(* IEC 61131-3 sources: daoli-st-library/DL_Device (part 33) *)

(* ---- FB_DL_ThreePointValve.st ---- *)
(*==============================================================================
 * 组件名称 (Component)  : FB_DL_ThreePointValve
 * 所属子库 (Sublibrary) : DL_Device
 * 当前版本 (Version)    : 1.0.1
 * 兼容性   (Platform)   : CODESYS 3.5 / TwinCAT 3 / 汇川 InoProShop / Machine Expert
 *                         仅依赖 Standard.library（TON / R_TRIG），零厂商方言
 * 分类     (Category)   : 设备执行器功能块（Function Block，实现 I_DL_MotorizedValve）
 * 功能简述 (Function)   : 三点浮点式电动调节阀控制器。开/关双脉冲输出；
 *                         行程时间积分自动估算开度（TON 计时段 ET 折算，
 *                         量纲推导见段 4 注释）；全开/全关限位双保险保护
 *                         （限位锚定 + 无限位端点拒绝）；限位互斥与估算-
 *                         限位一致性监视；双向指令互斥；首扫按限位状态
 *                         推断初值（R19 范式，bTrack 强制重同步）；状态机
 *                         E_DL_MotorValveState + CASE + ELSE 兜底。
 * 接口实现 (Implements) : I_DL_MotorizedValve。接口 OUT 列同名成员
 *                         （eState/fPosEstimate/bLimOpen/bLimClosed/
 *                         bFault/uErrorId）按 R22 以只读 PROPERTY GET 承载
 *                         （内部镜像同源；fPosEstimate 为 OUT 引脚、
 *                         bLimOpen/bLimClosed 为 IN 引脚与接口属性双形式
 *                         暴露，沿用库级既有先例），非接口成员 bOpenPulse/
 *                         bClosePulse/bOpened/bClosed/uTravelCount 保留
 *                         VAR_OUTPUT；方法 CmdOpen/CmdClose/CmdStop/
 *                         CmdReset 全部在本文件尾部落地。
 * 开源溯源 (Origin)     : 来源标签 lbp-basic-process / lbp-device
 *                         （RAW_NOTES_R6 S-1 + S-5：三点浮点式电动阀的开/
 *                         关脉冲控制、行程时间开度积分估算、端点限位双
 *                         保险等行业公知工程惯例，公开教学资料，仅借鉴
 *                         通用工程语义；状态机、积分实现、故障码按本库
 *                         红线独立设计，clean-room 未复制源码）。
 * 红线自检 (Redline)    : R1 零全局变量表/外部变量引用 ✓｜R2 零物理 IO 地址 ✓
 *                         R3 纯 IEC 61131-3 ✓｜R4 防除零/防越界/浮点容差
 *                         比较 ✓｜R5 全变量中英双语同行注释 ✓
 *                         R6 ENUM+CASE+ELSE ✓｜R7 四个定时器/边缘实例主体
 *                         最前部无条件刷新 ✓
 * 公约遵循 (Convention) : 0.1/R19 本块为事件型 + 连续估算混合组件：开度
 *                         积分为连续量，设 bInit 首扫（初值 FALSE，同步后
 *                         置 TRUE），判据唯一合法范式 IF bTrack OR (NOT
 *                         bInit)；bTrack 引脚供上层运行中途强制重同步。
 *                         0.7 故障码段位 16#0003_xxxx：【故障级】0003_0270
 *                         行程估算失准 / 0003_0271 双限位冲突 / 0003_0272
 *                         非法状态，R15 锁存仅复位可清；【信息级】
 *                         0003_0110 端点指令拒绝 / 0003_0111 双向指令冲突
 *                         （瞬时型每拍重算，0.15；不进 bFault）。
 * 偏离留档 (Deviation)  : 依 R11 头注释留档，共 3 条：
 *                         ① 信息级码：规格原分配 0003_0107/0108，经与子库
 *                           VERSION.md 故障码表核对，R5 已占用 0102~0104，
 *                           且 0106~0109 已由本轮变频器/模拟量阀块顺延占用
 *                           （0105 经终审裁定空置：重启抑制拒绝统一沿用
 *                           DolMotor 既有语义码位 0208），依公约 0.7 冲突
 *                           顺延为 0003_0110/0111。
 *                         ② 开度积分：规格原文"每拍按 fDt 增量累加"需周期
 *                           时间注入或时钟基准（与公约 0.9 冲突）；本实现
 *                           改用 TON 计时段 ET 累计行程时间折算：
 *                           fPosEstimate = 锚点 + 100 × ET[ms] / 行程时间[ms]
 *                           （量纲推导：无量纲比值 × 100% = [%]），等价
 *                           消除逐拍折算误差且零时钟依赖。
 *                         ③ bOpened/bClosed 的估算近似判据取固定 1% 吸附带
 *                           （限位优先，无限位场景估算到端点 1% 带内即视为
 *                           确认），规格未定值，现场可按需整定行程时间。
 * 修订历史 (Revision)   :
 *   2026-11-15  v1.0.0  首版入库（R6 轮 · DL_Device 阀门/驱动族深化）
 *   2026-11-15  v1.0.1  终审注释级修订：头注释偏离①码位占位表述与终审裁定
 *                       对齐（0105 空置、重启抑制拒绝归一 DolMotor 0208）。
 *                       逻辑零变更。已知诊断口径观察项（不改码）：uTravelCount
 *                       在上电首扫若全关限位已压住会即计 +1（限位态计数），
 *                       与 R4 PwmDutyController 首周期计数偏差同类，±1 口径。
 *============================================================================*)
FUNCTION_BLOCK FB_DL_ThreePointValve IMPLEMENTS I_DL_MotorizedValve
VAR_INPUT
    bCmdOpen     : BOOL;            // 开阀指令（Open command），电平生效 / Open command, level effective
    bCmdClose    : BOOL;            // 关阀指令（Close command），电平生效；与开同拍为真 → 停止 + 信息级 / Close command, conflict with open stops with info code
    bLimOpen     : BOOL;            // 全开限位开关（Open limit switch），TRUE=已到全开端点 / Open limit switch, TRUE = at fully-open endpoint
    bLimClosed   : BOOL;            // 全关限位开关（Closed limit switch），TRUE=已到全关端点 / Closed limit switch, TRUE = at fully-closed endpoint
    tStrokeOpen  : TIME := T#60S;   // 全行程开启时间（Full open stroke time），现场实测注入 / Full-open stroke time, field-measured
    tStrokeClose : TIME := T#60S;   // 全行程关闭时间（Full close stroke time），现场实测注入 / Full-close stroke time, field-measured
    fEstimateTol : REAL := 10.0;    // 估算-限位一致性容差（Estimate tolerance）[%]，默认 10.0 / Estimate-vs-limit consistency tolerance [%]
    bEnable      : BOOL;            // 允许动作联锁（Motion interlock），TRUE=允许发脉冲 / Motion interlock, TRUE = pulses allowed
    bReset       : BOOL;            // 故障复位（Fault reset），上升沿生效 / Fault reset, rising edge effective
    bTrack       : BOOL;            // 跟踪重同步（Track resync），TRUE 拍按限位状态重推初值（R19）/ Track resync re-infers initial estimate from limits
END_VAR

VAR_OUTPUT
    bOpenPulse   : BOOL;            // 开阀脉冲输出（Open pulse output）/ Open pulse output
    bClosePulse  : BOOL;            // 关阀脉冲输出（Close pulse output）/ Close pulse output
    fPosEstimate : REAL;            // 估算开度（Estimated position）[%]，0~100，行程时间积分（R20：量纲 [%]）/ Estimated position [%], stroke-time integration
    bOpened      : BOOL;            // 全开确认（Fully opened），限位优先 / Fully opened, limit switch has priority
    bClosed      : BOOL;            // 全关确认（Fully closed），限位优先 / Fully closed, limit switch has priority
    uTravelCount : UDINT;           // 全行程计数（Travel count），全关确认沿 +1 / Travel count, incremented on closed-confirmation edge
END_VAR

VAR
    _eState        : E_DL_MotorValveState := E_DL_MotorValveState.eIdle; // 内部状态机步序（Internal state step），外部经属性只读 / Internal state, read-only via property
    _bInit         : BOOL := FALSE; // 首扫初始化标志（First-scan init flag），R19 范式判据成员 / R19 paradigm member
    _bFaultLatch   : BOOL;          // 故障锁存标志（Fault latch flag），仅复位清除 / Fault latch flag, cleared only by reset
    _uErrorIdInt   : UDINT;         // 故障级码内部寄存（Internal fault-code register）/ Internal fault-level code register
    _uInfoCode     : UDINT;         // 本拍信息级码（Info code this cycle），瞬时型每拍重算（0.15）/ Transient info code recomputed each cycle
    _fAnchor       : REAL := 50.0;  // 积分锚点（Integration anchor）[%]，脉冲静止期与估算值同步 / Integration anchor [%], synced with estimate when idle
    _fEstInt       : REAL := 50.0;  // 估算开度内部寄存（Internal estimate register）[%] / Internal estimate register [%]
    _bPendOpen     : BOOL;          // 方法开阀保持锁存（Method open hold latch）/ Method open hold latch
    _bPendClose    : BOOL;          // 方法关阀保持锁存（Method close hold latch）/ Method close hold latch
    _bPendStop     : BOOL;          // 方法停止请求（Method stop request），由 CmdStop 置位 / Method stop request set by CmdStop
    _bPendReset    : BOOL;          // 方法复位请求（Method reset request），由 CmdReset 置位 / Method reset request set by CmdReset
    _bOpenReq      : BOOL;          // 合成开阀指令（Merged open command），引脚 OR 方法锁存 / Merged open command, pin OR method latch
    _bCloseReq     : BOOL;          // 合成关阀指令（Merged close command），引脚 OR 方法锁存 / Merged close command, pin OR method latch
    _bConflict     : BOOL;          // 双向同拍冲突（Open/close conflict this cycle）/ Open-close conflict flag
    _bOpenAtEnd    : BOOL;          // 开端点到达（Open endpoint reached），限位或估算判据 / Open endpoint reached by limit or estimate
    _bCloseAtEnd   : BOOL;          // 关端点到达（Close endpoint reached），限位或估算判据 / Close endpoint reached by limit or estimate
    _fTolEff       : REAL := 10.0;  // 防御后一致性容差（Sanitized tolerance）[%] / Sanitized consistency tolerance
    _tStrokeOpenEff  : TIME := T#60S; // 防御后开启行程时间（Sanitized open stroke time），非正值回退默认 / Sanitized open stroke time, non-positive falls back
    _tStrokeCloseEff : TIME := T#60S; // 防御后关闭行程时间（Sanitized close stroke time），非正值回退默认 / Sanitized close stroke time, non-positive falls back
    _bClosedInt    : BOOL;          // 全关确认内部镜像（Internal closed-confirmation mirror），喂计数边缘实例 / Internal closed mirror feeding count edge
    _bLimOpenMir   : BOOL;          // 全开限位内部镜像（Internal open-limit mirror），供属性读取 / Internal open-limit mirror for property exposure
    _bLimClosedMir : BOOL;          // 全关限位内部镜像（Internal closed-limit mirror），供属性读取 / Internal closed-limit mirror for property exposure
    _fbTrigReset   : R_TRIG;        // 引脚复位上升沿（Pin reset edge）/ Pin reset rising edge
    _fbTrigTravel  : R_TRIG;        // 全关确认计数上升沿（Travel count edge）/ Rising edge on closed confirmation for counting
    _fbTonOpenET   : TON;           // 开阀计时段定时器（Open timing segment timer），ET 供积分折算 / Open segment timer, ET feeds integration
    _fbTonCloseET  : TON;           // 关阀计时段定时器（Close timing segment timer），ET 供积分折算 / Close segment timer, ET feeds integration
END_VAR

METHOD CmdOpen : BOOL
VAR_INPUT
END_VAR
IF _bFaultLatch OR (_eState = E_DL_MotorValveState.eFault) THEN
    CmdOpen := FALSE;         // 故障态拒绝（Rejected in fault state）
    _bPendClose := FALSE;     // 清反向残留锁存（Clear stale reverse latch）
ELSE
    _bPendOpen := TRUE;       // 登记开阀保持锁存（Register open hold latch）
    _bPendClose := FALSE;     // 互斥注销关阀锁存（Cancel opposite close latch）
    CmdOpen := TRUE;          // 受理成功（Accepted）
END_IF

(*------------------------------------------------------------------------------
 * 方法: CmdClose —— 关阀指令（受理为保持锁存）。故障态一律拒绝返回 FALSE。
 *      Method CmdClose - close command held as latch, rejected with FALSE in fault.
 *------------------------------------------------------------------------------*)
    END_METHOD

METHOD CmdClose : BOOL
VAR_INPUT
END_VAR
IF _bFaultLatch OR (_eState = E_DL_MotorValveState.eFault) THEN
    CmdClose := FALSE;        // 故障态拒绝（Rejected in fault state）
    _bPendOpen := FALSE;      // 清反向残留锁存（Clear stale reverse latch）
ELSE
    _bPendClose := TRUE;      // 登记关阀保持锁存（Register close hold latch）
    _bPendOpen := FALSE;      // 互斥注销开阀锁存（Cancel opposite open latch）
    CmdClose := TRUE;         // 受理成功（Accepted）
END_IF

(*------------------------------------------------------------------------------
 * 方法: CmdStop —— 双脉冲全断保持当前位置。无条件受理。
 *      Method CmdStop - both pulses off and hold position, unconditionally accepted.
 *------------------------------------------------------------------------------*)
    END_METHOD

METHOD CmdStop : BOOL
VAR_INPUT
END_VAR
_bPendOpen  := FALSE;         // 注销开阀锁存（Cancel open latch）
_bPendClose := FALSE;         // 注销关阀锁存（Cancel close latch）
_bPendStop  := TRUE;          // 登记停止请求，主体状态机消化（Register stop request, consumed by body）
CmdStop := TRUE;              // 无条件受理（Unconditionally accepted）

(*------------------------------------------------------------------------------
 * 方法: CmdReset —— 复位故障，返回是否可复位（存在锁存故障时为 TRUE）。
 *      Method CmdReset - reset fault, returns TRUE only when a latch exists.
 *------------------------------------------------------------------------------*)
    END_METHOD

METHOD CmdReset : BOOL
VAR_INPUT
END_VAR
IF _bFaultLatch OR (_eState = E_DL_MotorValveState.eFault) THEN
    _bPendReset := TRUE;      // 登记复位请求，主体状态机消化（Register reset request, consumed by body）
    CmdReset := TRUE;         // 可复位（Resettable）
ELSE
    CmdReset := FALSE;        // 无故障可复位（Nothing to reset）
END_IF

(*------------------------------------------------------------------------------
 * 属性: eState（GET）—— 当前状态机状态只读视图。
 *      Property eState (GET) - read-only view of the current state machine state.
 *------------------------------------------------------------------------------*)
    END_METHOD

// ============================================================================
// 段 1｜定时器与边缘检测实例无条件周期刷新（R7：严禁置于 IF/CASE 分支内）
//      Unconditional per-cycle refresh of all timer and edge instances (R7)
// ============================================================================
_fbTrigReset(CLK := bReset);
_fbTonOpenET(IN := bOpenPulse, PT := _tStrokeOpenEff);   // 计时段随开阀脉冲累计（Segment ET accumulates with open pulse）
_fbTonCloseET(IN := bClosePulse, PT := _tStrokeCloseEff); // 计时段随关阀脉冲累计（Segment ET accumulates with close pulse）
_bClosedInt := bLimClosed OR (_fEstInt <= 1.0);           // 全关确认镜像（Closed-confirmation mirror, limit priority + 1% snap band）
_fbTrigTravel(CLK := _bClosedInt);
IF _fbTrigTravel.Q THEN
    uTravelCount := uTravelCount + 1;                     // 全行程计数 +1（Travel count +1 on closed confirmation）
END_IF

// ============================================================================
// 段 2｜首扫/跟踪初始化（R19 唯一合法范式：IF bTrack OR (NOT bInit)）
//      First-scan / track initialization (R19 sole legal paradigm)
// ============================================================================
IF bTrack OR (NOT _bInit) THEN
    IF bLimOpen THEN
        _fAnchor := 100.0;                // 限位推断：已全开（Inferred from limit: fully open）
    ELSIF bLimClosed THEN
        _fAnchor := 0.0;                  // 限位推断：已全关（Inferred from limit: fully closed）
    ELSE
        _fAnchor := 50.0;                 // 无限位信息：中位兜底（No limit info: mid-position fallback）
    END_IF
    _fEstInt := _fAnchor;                 // 估算值与锚点同步（Estimate synced with anchor）
    _bInit  := TRUE;                      // 初始化完成（Initialization done）
END_IF

// ============================================================================
// 段 3｜参数防御（0.8）+ 指令合成与冲突判定
//      Parameter sanitation (0.8) + command merge and conflict evaluation
// ============================================================================
_uInfoCode := 0;                          // 本拍信息级码先归零，事件分支重算（Info code preset zero, recomputed in branches）
_bLimOpenMir := bLimOpen;                 // 全开限位镜像刷新（Refresh open-limit mirror）
_bLimClosedMir := bLimClosed;             // 全关限位镜像刷新（Refresh closed-limit mirror）
_fTolEff := fEstimateTol;                 // 容差镜像（Tolerance mirror）
IF _fTolEff <> _fTolEff THEN              // 非数自比检测（NaN self-compare test）
    _fTolEff := 10.0;                     // 回落默认容差（Fallback to default tolerance）
END_IF
IF _fTolEff < 0.0 THEN
    _fTolEff := ABS(_fTolEff);            // 负容差取绝对值（Negative tolerance made absolute）
END_IF
_tStrokeOpenEff := tStrokeOpen;           // 开启行程时间镜像（Open stroke time mirror）
IF _tStrokeOpenEff <= T#0S THEN
    _tStrokeOpenEff := T#60S;             // 非正值回退默认，防积分除零（Non-positive falls back, divide-by-zero guard）
END_IF
_tStrokeCloseEff := tStrokeClose;         // 关闭行程时间镜像（Close stroke time mirror）
IF _tStrokeCloseEff <= T#0S THEN
    _tStrokeCloseEff := T#60S;            // 非正值回退默认，防积分除零（Non-positive falls back, divide-by-zero guard）
END_IF

_bOpenReq := bCmdOpen OR _bPendOpen;      // 合成开阀指令（Merged open command）
_bCloseReq := bCmdClose OR _bPendClose;   // 合成关阀指令（Merged close command）
_bConflict := _bOpenReq AND _bCloseReq;   // 双向同拍冲突（Same-cycle conflict）
IF _bConflict THEN
    _uInfoCode := 16#0003_0111;           // 0003_0111 双向指令冲突【信息级】/ Open-close conflict, info level
END_IF
_bOpenAtEnd := bLimOpen OR (_fEstInt >= 100.0);    // 开端点判据（Open endpoint test）
_bCloseAtEnd := bLimClosed OR (_fEstInt <= 0.0);   // 关端点判据（Close endpoint test）

// ============================================================================
// 段 4｜开度积分（换算式：估算 = 锚点 + 100 × 计时段ET[ms] / 行程时间[ms]，
//       无量纲比值 × 100% → 量纲 [%]，R20；钳位 [0,100]；脉冲静止期锚点
//       与估算同步）
//      Position integration (see conversion formula above; clamped [0,100];
//      anchor synced with estimate while pulses idle)
// ============================================================================
IF bLimOpen THEN
    _fAnchor := 100.0;                    // 限位锚定：全开（Limit anchor: fully open）
    _fEstInt := 100.0;
ELSIF bLimClosed THEN
    _fAnchor := 0.0;                      // 限位锚定：全关（Limit anchor: fully closed）
    _fEstInt := 0.0;
ELSIF bOpenPulse THEN
    _fEstInt := _fAnchor + (100.0 * (TIME_TO_REAL(_fbTonOpenET.ET) / TIME_TO_REAL(_tStrokeOpenEff))); // 开向积分（Open-direction integration, divisor proven positive）
    IF _fEstInt > 100.0 THEN
        _fEstInt := 100.0;                // 上限钳位（Clamped to high bound）
    END_IF
ELSIF bClosePulse THEN
    _fEstInt := _fAnchor - (100.0 * (TIME_TO_REAL(_fbTonCloseET.ET) / TIME_TO_REAL(_tStrokeCloseEff))); // 关向积分（Close-direction integration, divisor proven positive）
    IF _fEstInt < 0.0 THEN
        _fEstInt := 0.0;                  // 下限钳位（Clamped to low bound）
    END_IF
ELSE
    _fAnchor := _fEstInt;                 // 脉冲静止期：锚点与估算同步（Pulses idle: anchor synced with estimate）
END_IF

// ============================================================================
// 段 5｜限位与估算一致性全局监视（优先级最高，故障级锁存）
//      Limit and estimate consistency global monitor (highest priority)
// ============================================================================
IF bLimOpen AND bLimClosed THEN
    _bFaultLatch := TRUE;                 // 双限位冲突锁存（Dual-limit conflict latch）
    _uErrorIdInt := 16#0003_0271;         // 0003_0271 双限位冲突（物理不可能）【故障级】/ Dual-limit conflict, fault level
    _eState      := E_DL_MotorValveState.eFault; // 强制故障态（Force fault state）
ELSIF bLimClosed AND (_fEstInt > _fTolEff) THEN
    _bFaultLatch := TRUE;                 // 估算失准锁存（Estimate mismatch latch）
    _uErrorIdInt := 16#0003_0270;         // 0003_0270 行程估算失准（估算与限位矛盾超容差）【故障级】/ Estimate mismatch beyond tolerance, fault level
    _eState      := E_DL_MotorValveState.eFault;
ELSIF bLimOpen AND (_fEstInt < (100.0 - _fTolEff)) THEN
    _bFaultLatch := TRUE;                 // 估算失准锁存（Estimate mismatch latch）
    _uErrorIdInt := 16#0003_0270;         // 0003_0270 行程估算失准【故障级】/ Estimate mismatch beyond tolerance, fault level
    _eState      := E_DL_MotorValveState.eFault;
END_IF

// ============================================================================
// 段 6｜核心状态机（ENUM + CASE，含 ELSE 非法状态兜底）
//      Core state machine (ENUM + CASE with ELSE illegal-state fallback)
// ============================================================================
IF _bFaultLatch OR (_eState = E_DL_MotorValveState.eFault) THEN
    CASE _eState OF
        E_DL_MotorValveState.eFault: // 故障锁存态：清空全部请求，仅复位可退出
            _bPendOpen  := FALSE;             // 清方法锁存（Clear method latches）
            _bPendClose := FALSE;
            _bPendStop  := FALSE;
            IF _bPendReset OR _fbTrigReset.Q THEN
                _bPendReset  := FALSE;        // 消费复位请求（Consume reset request）
                _bFaultLatch := FALSE;        // 解除锁存（Release latch）
                _uErrorIdInt := 0;            // 故障码清零（Error code cleared）
                _fAnchor     := _fEstInt;     // 锚点与估算重同步（Anchor re-synced with estimate）
                _eState      := E_DL_MotorValveState.eIdle; // 回空闲态（Back to idle）
            END_IF
        ELSE // 锁存标志与状态不一致兜底：强制同步进故障态（Latch/state mismatch fallback）
            _eState := E_DL_MotorValveState.eFault;
    END_CASE
ELSE
    CASE _eState OF

        E_DL_MotorValveState.eIdle: // 空闲稳态：双脉冲全断
            IF _bPendStop THEN
                _bPendStop := FALSE;          // 消化停止请求（Absorb stop request）
            END_IF
            IF bLimOpen THEN
                _fAnchor := 100.0;            // 限位同步锚点（Sync anchor with limit）
                _fEstInt := 100.0;
                _eState  := E_DL_MotorValveState.eOpened;
            ELSIF bLimClosed THEN
                _fAnchor := 0.0;              // 限位同步锚点（Sync anchor with limit）
                _fEstInt := 0.0;
                _eState  := E_DL_MotorValveState.eClosed;
            ELSIF _bConflict THEN
                // 双向冲突：安全侧不动，信息级已在段 3 置码（Conflict: hold, info code set in section 3）
            ELSIF _bOpenReq AND (NOT _bOpenAtEnd) THEN
                _eState := E_DL_MotorValveState.eOpening; // 受理开阀（Accept open）
            ELSIF _bCloseReq AND (NOT _bCloseAtEnd) THEN
                _eState := E_DL_MotorValveState.eClosing; // 受理关阀（Accept close）
            ELSIF (_bOpenReq AND _bOpenAtEnd) OR (_bCloseReq AND _bCloseAtEnd) THEN
                _uInfoCode := 16#0003_0110;   // 0003_0110 端点指令拒绝【信息级】/ Endpoint command refused, info level
            END_IF

        E_DL_MotorValveState.eOpening: // 开阀中：开阀脉冲输出
            IF bLimOpen THEN
                _fAnchor := 100.0;            // 限位锚定双保险①（Limit anchor, protection layer 1）
                _fEstInt := 100.0;
                _eState  := E_DL_MotorValveState.eOpened;
            ELSIF (NOT _bOpenReq) OR _bConflict OR _bPendStop THEN
                _bPendStop := FALSE;          // 消化停止请求（Absorb stop request）
                _eState    := E_DL_MotorValveState.eIdle; // 指令撤除/冲突/停止：回空闲（Command dropped, conflict or stop: to idle）
            ELSIF _fEstInt >= 100.0 THEN
                _uInfoCode := 16#0003_0110;   // 0003_0110 端点指令拒绝（无限位端点双保险②）【信息级】/ Endpoint refused (no-limit protection layer 2), info level
                _eState    := E_DL_MotorValveState.eIdle;
            END_IF

        E_DL_MotorValveState.eClosing: // 关阀中：关阀脉冲输出
            IF bLimClosed THEN
                _fAnchor := 0.0;              // 限位锚定双保险①（Limit anchor, protection layer 1）
                _fEstInt := 0.0;
                _eState  := E_DL_MotorValveState.eClosed;
            ELSIF (NOT _bCloseReq) OR _bConflict OR _bPendStop THEN
                _bPendStop := FALSE;          // 消化停止请求（Absorb stop request）
                _eState    := E_DL_MotorValveState.eIdle; // 指令撤除/冲突/停止：回空闲（Command dropped, conflict or stop: to idle）
            ELSIF _fEstInt <= 0.0 THEN
                _uInfoCode := 16#0003_0110;   // 0003_0110 端点指令拒绝（无限位端点双保险②）【信息级】/ Endpoint refused (no-limit protection layer 2), info level
                _eState    := E_DL_MotorValveState.eIdle;
            END_IF

        E_DL_MotorValveState.eOpened: // 全开确认稳态：限位优先
            IF NOT bLimOpen THEN
                _eState := E_DL_MotorValveState.eIdle; // 限位脱开回空闲（Limit dropped, to idle）
            ELSIF _bCloseReq AND (NOT _bCloseAtEnd) THEN
                _eState := E_DL_MotorValveState.eClosing; // 受理关阀（Accept close）
            ELSIF _bOpenReq THEN
                _uInfoCode := 16#0003_0110;   // 0003_0110 端点指令拒绝（限位确认端点）【信息级】/ Endpoint command refused at limit, info level
            END_IF

        E_DL_MotorValveState.eClosed: // 全关确认稳态：限位优先
            IF NOT bLimClosed THEN
                _eState := E_DL_MotorValveState.eIdle; // 限位脱开回空闲（Limit dropped, to idle）
            ELSIF _bOpenReq AND (NOT _bOpenAtEnd) THEN
                _eState := E_DL_MotorValveState.eOpening; // 受理开阀（Accept open）
            ELSIF _bCloseReq THEN
                _uInfoCode := 16#0003_0110;   // 0003_0110 端点指令拒绝（限位确认端点）【信息级】/ Endpoint command refused at limit, info level
            END_IF

        ELSE // 非法状态兜底：任何越界枚举值强制锁存故障（Illegal state fallback）
            _bFaultLatch := TRUE;             // 故障锁存（Fault latched）
            _uErrorIdInt := 16#0003_0272;     // 0003_0272 非法状态【故障级】/ Illegal state, fault level
            _eState      := E_DL_MotorValveState.eFault;
    END_CASE
END_IF

// ============================================================================
// 段 7｜脉冲输出推导 + 双脉冲互斥出口断言（硬约束：开/关脉冲恒不可同真）
//      Pulse output derivation + mutual exclusivity exit assertion
// ============================================================================
bOpenPulse  := (_eState = E_DL_MotorValveState.eOpening) AND _bOpenReq AND (NOT _bConflict)
               AND bEnable AND (NOT bLimOpen) AND (_fEstInt < 100.0); // 开阀脉冲使能条件链（Open pulse condition chain）
bClosePulse := (_eState = E_DL_MotorValveState.eClosing) AND _bCloseReq AND (NOT _bConflict)
               AND bEnable AND (NOT bLimClosed) AND (_fEstInt > 0.0); // 关阀脉冲使能条件链（Close pulse condition chain）
IF bOpenPulse AND bClosePulse THEN
    bOpenPulse  := FALSE;               // 断言对调：异常同真时双断保安全（Assertion fallback: cut both on impossible condition）
    bClosePulse := FALSE;
END_IF
IF (_eState = E_DL_MotorValveState.eFault) OR (_eState = E_DL_MotorValveState.eIdle)
   OR (_eState = E_DL_MotorValveState.eOpened) OR (_eState = E_DL_MotorValveState.eClosed) THEN
    bOpenPulse  := FALSE;               // 出口断言：非动作态脉冲必断（Assertion: pulses off in non-motion states）
    bClosePulse := FALSE;
END_IF
fPosEstimate := _fEstInt;               // 估算开度输出（Estimate output）
bOpened := bLimOpen OR (_fEstInt >= 99.0); // 全开确认：限位优先 + 1% 吸附带（Opened: limit priority + 1% snap band）
bClosed := bLimClosed OR (_fEstInt <= 1.0); // 全关确认：限位优先 + 1% 吸附带（Closed: limit priority + 1% snap band）

(*------------------------------------------------------------------------------
 * 方法: CmdOpen —— 开阀指令（受理为保持锁存）。故障态一律拒绝返回 FALSE。
 *      Method CmdOpen - open command held as latch, rejected with FALSE in fault.
 *------------------------------------------------------------------------------*)

PROPERTY eState : E_DL_MotorValveState
eState := _eState;            // 返回内部状态（Return internal state）

(*------------------------------------------------------------------------------
 * 属性: fPosEstimate（GET）—— 估算开度 [%]（行程时间积分）。
 *      Property fPosEstimate (GET) - estimated position [%] from stroke-time integration.
 *------------------------------------------------------------------------------*)
PROPERTY fPosEstimate : REAL
fPosEstimate := _fEstInt;     // 返回估算镜像（Return estimate mirror）

(*------------------------------------------------------------------------------
 * 属性: bLimOpen（GET）—— 全开限位反馈。
 *      Property bLimOpen (GET) - open limit switch feedback.
 *------------------------------------------------------------------------------*)
PROPERTY bLimOpen : BOOL
bLimOpen := _bLimOpenMir;     // 返回限位镜像（Return limit mirror）

(*------------------------------------------------------------------------------
 * 属性: bLimClosed（GET）—— 全关限位反馈。
 *      Property bLimClosed (GET) - closed limit switch feedback.
 *------------------------------------------------------------------------------*)
PROPERTY bLimClosed : BOOL
bLimClosed := _bLimClosedMir; // 返回限位镜像（Return limit mirror）

(*------------------------------------------------------------------------------
 * 属性: bFault（GET）—— 故障锁存指示（信息级码不置本位，0.2 公约）。
 *      Property bFault (GET) - fault latch indicator, info-level codes excluded.
 *------------------------------------------------------------------------------*)
PROPERTY bFault : BOOL
bFault := _bFaultLatch OR (_eState = E_DL_MotorValveState.eFault); // 显式排除信息级派生式（Explicit derived form excluding info codes）

(*------------------------------------------------------------------------------
 * 属性: uErrorId（GET）—— 末次事件码（故障级锁存优先；无故障时透出本拍
 *         信息级码，0.2/0.15 公约）。
 *      Property uErrorId (GET) - last event code (fault-level priority,
 *      transient info code shown otherwise).
 *------------------------------------------------------------------------------*)
PROPERTY uErrorId : UDINT
IF (_uErrorIdInt <> 0) OR (_eState = E_DL_MotorValveState.eFault) THEN
    uErrorId := _uErrorIdInt; // 故障级码优先透出（Fault-level code has priority）
ELSE
    uErrorId := _uInfoCode;   // 无故障时透出本拍信息级码（Transient info code when no fault）
END_IF
END_FUNCTION_BLOCK

(* ---- FB_DL_TwoSpeedMotor.st ---- *)
(*==============================================================================
 * 组件名称 (Component)  : FB_DL_TwoSpeedMotor
 * 所属子库 (Sublibrary) : DL_Device
 * 当前版本 (Version)    : 1.0.1
 * 兼容性   (Platform)   : CODESYS 3.5 / TwinCAT 3 / 汇川 InoProShop / Machine Expert
 *                         仅依赖 Standard.library（TON / R_TRIG），零厂商方言
 * 来源标签 (Source)     : t2-2-lbp（电机族 · 变极双速驱动，clean-room 编写）
 * 功能描述 (Function)   : 双绕组变极调速驱动：低速 / 高速选择 + 切换死区互锁
 *                         （低速断电 -> 死区窗内双绕组全断 -> 高速投入）+ 高速
 *                         禁止位（工艺联锁，优先于一切运行请求）+ 两方向接触器
 *                         反馈校验。死区窗内任一异侧反馈已出现即判绕组粘连故障
 *                         （锁存 + 安全侧断高速）；投入后反馈超时未到判校验失败。
 * 范式次源 (Paradigm)   : 命令-反馈范式参照 I_DL_MotorDriver 契约；星角切换安全
 *                         死区范式参照 FB_DL_StarDeltaMotor（互引声明，不复用实现、
 *                         不共享枚举——变极为双独立绕组，无星角三态）。
 * 配比约束 (R100)       : tFbTimeout > tDeadZone（反馈校验窗必须宽于死区窗，
 *                         否则死区未结束即误判反馈超时）。
 * 边界与语义披露 (Boundary disclosure) :
 *   1) 切换期间两绕组互斥硬闸：统一出口对 bOutLow / bOutHigh 再做 AND NOT 交叉
 *      硬闸，CASE 内任何路径都不可能产出双投（结构 + 出口双保险）。
 *   2) 死区窗内反馈校验（粘连判据）：命令已断侧的反馈若仍为 TRUE，判绕组粘连
 *      （机械/触点粘连），立即中止切换并锁存；高速粘连按安全侧断高速。
 *   3) 高速禁止位优先于一切运行请求：禁止位有效时高速请求被拒（信息级），运行中
 *      高速遇禁止位即时降速切换（不等待操作员）。
 *   4) 死区组态非法（<= T#0S）拒绝一切新切换，已运行的绕组保持（组态错误不停机，
 *      但故障级码必须可见，R191 显式声明）。
 *   5) 失能语义声明：bEnable = FALSE 时双绕组全断（安全侧），不冻结保持。
 * 故障码表 (Error codes) :
 *   16#0003_050B [故障级] 绕组粘连：死区窗内异侧反馈已出现，中止切换 + 锁存
 *                 反证：粘连拍输出与正常切换拍组合不同仅在于「反馈先行」，无码
 *                 则操作员只见切换中止不见根因。
 *   16#0003_050C [故障级] 反馈校验失败：投入命令已发而反馈超时未到，锁存 + 断高速
 *                 反证：校验失败与粘连状态输出组合不同（一为无反馈一为多反馈），
 *                 两因必须码位互异（R190）。
 *   16#0003_050D [故障级] 死区组态非法（<= T#0S），拒绝新切换 + 锁存
 *                 反证：拒绝切换与「无切换请求」输出组合相同，码位唯一可见。
 *   16#0003_0409 [信息级] 高速请求被禁止位拒绝（工艺联锁生效）
 *                 反证：请求被拒时电机保持低速，与「本来就选低速」输出组合相同，
 *                 无码则联锁生效事实不可观测。
 * 码位总账 (Code ledger) : 16#0003_050B / 050C / 050D 用 ｜ 16#0003_0409 用
 * 依赖     (Depends)    : 无 DL_ 内部依赖；Standard.library: TON / R_TRIG
 * 红线自检 (Redline)    : R1 ✓ 零全局变量与 VAR_EXTERNAL ｜ R2 ✓ 零 %I/%Q 物理地址
 *                         R3 ✓ 纯 IEC 61131-3 ｜ R4 ✓ 域闸 / 计数无涉 / 码位 R45 配对
 *                         R5 ✓ 全变量中英双语同行注释 ｜ R6 ✓ 六态 ENUM + CASE + ELSE 兜底
 *                         R7 ✓ 三沿三计时主体最前部无条件刷新
 * 修订历史 (Revision)   :
 *   2026-11-22  v1.0.0  首版入库（R68 构建轮 · 批 2 · 目标 10）
 *   2026-11-22  v1.0.1  终审就地修①：组态锁存解除路径可达化（原 bCfgLatch 全文件零清零 -> 双绕组永久双断）
 *============================================================================*)

(*-----------------------------------------------------------------------------
 * 枚举: E_DL_TwoSpeedState（归属 DL_Device，与 FB_DL_TwoSpeedMotor 同文件）
 *----------------------------------------------------------------------------*)
TYPE E_DL_TwoSpeedState :
(
    eIdle    := 0,    // 停机：双绕组全断 / Stopped, both windings off
    eRunLow  := 10,   // 低速运行：低速绕组投入 / Low speed, low winding on
    eSwUp    := 20,   // 升速切换：死区窗内双绕组全断 / Speed-up transition, dead zone
    eRunHigh := 30,   // 高速运行：高速绕组投入 / High speed, high winding on
    eSwDown  := 40,   // 降速切换：死区窗内双绕组全断 / Speed-down transition, dead zone
    eFault   := 99    // 粘连 / 校验故障锁存：双绕组全断 / Latched fault, both off
);
END_TYPE

(*==============================================================================
 * 功能块: FB_DL_TwoSpeedMotor
 * 调用约定: 每个扫描周期无条件调用一次。
 *============================================================================*)
FUNCTION_BLOCK FB_DL_TwoSpeedMotor
VAR_INPUT
    bStartCmd   : BOOL;                  // 运行命令（电平）/ Run command, level
    bStopCmd    : BOOL;                  // 停止命令（电平，优先）/ Stop command, level, priority
    bHighReq    : BOOL;                  // 速度选择：TRUE = 高速请求 / Speed select, TRUE high speed
    bHighInhibit: BOOL;                  // 高速禁止位（工艺联锁）/ High speed inhibit, process interlock
    bFbLow      : BOOL;                  // 低速接触器反馈 / Low speed contactor feedback
    bFbHigh     : BOOL;                  // 高速接触器反馈 / High speed contactor feedback
    tDeadZone   : TIME := T#2S;          // 绕组切换死区窗 [s]，<= T#0S 组态非法 / Dead zone window [s]
    tFbTimeout  : TIME := T#3S;          // 反馈校验窗 [s]，须 > tDeadZone / Feedback verify window [s]
    bEnable     : BOOL := TRUE;          // 使能（FALSE 双绕组全断）/ Enable, FALSE cuts both
    bReset      : BOOL;                  // 上升沿：清除粘连 / 校验 / 组态锁存 / Rising edge: clear latches
END_VAR
VAR_OUTPUT
    bOutLow    : BOOL;                  // 低速绕组输出（经互斥硬闸）/ Low winding output, hard-gated
    bOutHigh   : BOOL;                  // 高速绕组输出（经互斥硬闸）/ High winding output, hard-gated
    bSwitching : BOOL;                  // 切换（死区窗）进行中 / Transition dead zone in progress
    bAdhesion  : BOOL;                  // 绕组粘连锁存 / Winding adhesion latched
    bFbFail    : BOOL;                  // 反馈校验失败锁存 / Feedback verify failed latched
    bError     : BOOL;                  // 故障标志（锁存类归并）/ Fault flag, latched class merged
    uErrorId   : UDINT;                 // 故障码，0 = 无故障 / Error code, 0 = none
    eState     : E_DL_TwoSpeedState;    // 当前状态（供 HMI 诊断）/ Current state for HMI diagnosis
END_VAR
VAR
    fbTrigReset  : R_TRIG;              // 复位沿检测实例 / Reset edge detector
    tonDead      : TON;                 // 切换死区窗计时实例 / Dead zone timer
    tonFbLow     : TON;                 // 低速反馈校验计时实例 / Low feedback verify timer
    tonFbHigh    : TON;                 // 高速反馈校验计时实例 / High feedback verify timer
    eStateInt    : E_DL_TwoSpeedState;  // 主状态机内部当前态 / Internal state machine state
    bOutLowInt   : BOOL;                // 低速输出内部副本（出口前未闸）/ Internal low output, pre-gate
    bOutHighInt  : BOOL;                // 高速输出内部副本（出口前未闸）/ Internal high output, pre-gate
    bDeadRun     : BOOL;                // 死区窗计时进行中 / Dead zone timing active
    bFbWaitLow   : BOOL;                // 低速反馈待达（投入后未反馈）/ Low feedback pending
    bFbWaitHigh  : BOOL;                // 高速反馈待达 / High feedback pending
    bAdhesionInt : BOOL;                // 粘锁存内部副本 / Internal adhesion latch
    bFbFailInt   : BOOL;                // 校验失败锁存内部副本 / Internal verify-fail latch
    bCfgLatch    : BOOL;                // 死区组态锁存（复位沿清除）/ Dead-zone config latch
    bCfgBad      : BOOL;                // 本拍死区组态非法 / Dead-zone config illegal this scan
    bHighRefused : BOOL;                // 高速请求被禁脉冲内部副本（单拍）/ Internal high-refused pulse
    bErrorInt    : BOOL;                // 本拍故障置位累加（出口归并）/ Fault set accumulator
    bFirstScan   : BOOL := TRUE;        // 上电首扫标志 / First-scan flag
END_VAR

(*------------------------------------------------------------------------------
 * 段 1｜无条件刷新区（红线 R7）：一沿三计时全部位于主体最前部
 *      Unconditional refresh: one edge and three timers at the very top
 *-----------------------------------------------------------------------------*)
fbTrigReset(CLK := bReset);

bFbWaitLow  := (eStateInt = E_DL_TwoSpeedState.eRunLow)  AND (NOT bFbLow);
bFbWaitHigh := (eStateInt = E_DL_TwoSpeedState.eRunHigh) AND (NOT bFbHigh);

tonDead(IN := bDeadRun, PT := tDeadZone);
tonFbLow(IN := bFbWaitLow, PT := tFbTimeout);
tonFbHigh(IN := bFbWaitHigh, PT := tFbTimeout);

(*------------------------------------------------------------------------------
 * 段 2｜上电首扫：双绕组全断落安全侧
 *      First-scan init: both windings to the safe off side
 *-----------------------------------------------------------------------------*)
IF bFirstScan THEN
    eStateInt   := E_DL_TwoSpeedState.eIdle;
    bOutLowInt  := FALSE;
    bOutHighInt := FALSE;
    bFirstScan  := FALSE;
END_IF

(*------------------------------------------------------------------------------
 * 段 3｜每拍预清（FB32-1）：单拍标志，禁入锁存 / 快照
 *      Per-scan preset: single-scan flags only
 *-----------------------------------------------------------------------------*)
bErrorInt    := FALSE;
bHighRefused := FALSE;

(*------------------------------------------------------------------------------
 * 段 4｜组态域闸（R151）+ 配比复检：死区 <= T#0S 拒绝新切换，运行绕组保持
 *      Config gate and ratio re-check: bad dead zone refuses new transitions
 *      解除路径（R152 自证）：复位沿 AND 死区组态已改对
 *-----------------------------------------------------------------------------*)
bCfgBad := (tDeadZone <= T#0S);

IF bCfgBad THEN
    bCfgLatch := TRUE;
    uErrorId  := 16#0003_050D;   // 故障级：死区组态非法 / Fault: dead zone config illegal
    bErrorInt := TRUE;
END_IF

(* 终审就地修 v1.0.1（R68）：解除路径（R152 自证可达）——复位沿 AND 组态非法条件
 * 全部消失即清锁存。原实现把锁存清零只写在 eFault 相分支，而组态闸置锁存后
 * 并不迁相至 eFault（只回 eIdle / 驻留），eFault 相不可达 -> 锁存永不可解，
 * 组件保护/监视功能一次性永久失效直至 PLC 重启（终审两式①）。
 * Clear path made provably reachable: reset edge with the illegal config gone. *)
IF fbTrigReset.Q AND (NOT bCfgBad) THEN
    bCfgLatch := FALSE;          // 锁存解除 / Latch cleared
    uErrorId  := 16#0000_0000;   // 码位随解除归零 / Code cleared with the latch
END_IF

(*------------------------------------------------------------------------------
 * 段 5｜主状态机（红线 R6）：ENUM + CASE + ELSE 兜底
 *      Main state machine with the mandatory ELSE fallback
 *-----------------------------------------------------------------------------*)
CASE eStateInt OF

    E_DL_TwoSpeedState.eIdle:
        IF (NOT bEnable) OR bStopCmd OR bCfgLatch THEN
            bOutLowInt  := FALSE;    // 双断驻留 / Both-off dwell
            bOutHighInt := FALSE;
        ELSIF bStartCmd THEN
            IF bHighReq AND bHighInhibit THEN
                bHighRefused := TRUE;    // 高速请求被禁止位拒绝（信息级）/ High refused by inhibit
                uErrorId     := 16#0003_0409;
                bOutLowInt   := TRUE;    // 抑制优先：按低速受理 / Inhibit wins: start low
                bOutHighInt  := FALSE;
                eStateInt    := E_DL_TwoSpeedState.eRunLow;
            ELSIF bHighReq THEN
                bOutLowInt  := FALSE;    // 高速直投：先断后投死区窗 / High direct: dead zone first
                bOutHighInt := FALSE;
                bDeadRun    := TRUE;
                eStateInt   := E_DL_TwoSpeedState.eSwUp;
            ELSE
                bOutLowInt  := TRUE;     // 低速直投（无死区需求）/ Low direct, no dead zone needed
                bOutHighInt := FALSE;
                eStateInt   := E_DL_TwoSpeedState.eRunLow;
            END_IF
        END_IF

    E_DL_TwoSpeedState.eRunLow:
        IF (NOT bEnable) OR bStopCmd THEN
            bOutLowInt  := FALSE;    // 停机双断 / Stop, both off
            bOutHighInt := FALSE;
            eStateInt   := E_DL_TwoSpeedState.eIdle;
        ELSIF bHighReq AND bHighInhibit THEN
            bHighRefused := TRUE;    // 禁止位拒高速（信息级，保持低速）/ High refused, keep low
            uErrorId     := 16#0003_0409;
        ELSIF bHighReq AND (NOT bCfgLatch) THEN
            bOutLowInt  := FALSE;    // 升速切换：先断低速 / Speed-up: drop low first
            bDeadRun    := TRUE;
            eStateInt   := E_DL_TwoSpeedState.eSwUp;
        END_IF

    E_DL_TwoSpeedState.eSwUp:
        (* 死区窗（升速）：双绕组全断；异侧反馈出现即粘连；窗满投高速 *)
        (* Dead zone up: both off; early feedback means adhesion; commit at window full *)
        IF (NOT bEnable) OR bStopCmd THEN
            bOutLowInt  := FALSE;    // 中止切换双断 / Abort, both off
            bOutHighInt := FALSE;
            bDeadRun    := FALSE;
            eStateInt   := E_DL_TwoSpeedState.eIdle;
        ELSIF bFbHigh OR bFbLow THEN
            bAdhesionInt := TRUE;    // 死区内反馈先行 = 绕组粘连 / Early feedback = adhesion
            uErrorId     := 16#0003_050B;
            bErrorInt    := TRUE;
            bOutHighInt  := FALSE;   // 安全侧断高速（本相本就全断，显式再声明）/ High cut on safe side
            bDeadRun     := FALSE;
            eStateInt    := E_DL_TwoSpeedState.eFault;
        ELSIF tonDead.Q THEN
            bOutHighInt := TRUE;     // 窗满投高速 / Window full, high on
            bDeadRun    := FALSE;
            eStateInt   := E_DL_TwoSpeedState.eRunHigh;
        END_IF

    E_DL_TwoSpeedState.eRunHigh:
        IF (NOT bEnable) OR bStopCmd THEN
            bOutLowInt  := FALSE;    // 停机双断 / Stop, both off
            bOutHighInt := FALSE;
            eStateInt   := E_DL_TwoSpeedState.eIdle;
        ELSIF bHighInhibit OR (NOT bHighReq) THEN
            bOutHighInt := FALSE;    // 禁止位优先 / 请求撤销：降速切换 / Inhibit or request gone: down-switch
            bDeadRun    := TRUE;
            eStateInt   := E_DL_TwoSpeedState.eSwDown;
        END_IF

    E_DL_TwoSpeedState.eSwDown:
        (* 死区窗（降速）：双绕组全断；异侧反馈出现即粘连；窗满投低速 *)
        (* Dead zone down: both off; early feedback means adhesion; commit low *)
        IF (NOT bEnable) OR bStopCmd THEN
            bOutLowInt  := FALSE;
            bOutHighInt := FALSE;
            bDeadRun    := FALSE;
            eStateInt   := E_DL_TwoSpeedState.eIdle;
        ELSIF bFbHigh OR bFbLow THEN
            bAdhesionInt := TRUE;    // 死区内反馈先行 = 绕组粘连 / Early feedback = adhesion
            uErrorId     := 16#0003_050B;
            bErrorInt    := TRUE;
            bOutHighInt  := FALSE;   // 安全侧断高速 / High cut on safe side
            bDeadRun     := FALSE;
            eStateInt    := E_DL_TwoSpeedState.eFault;
        ELSIF tonDead.Q THEN
            bOutLowInt := TRUE;      // 窗满投低速 / Window full, low on
            bDeadRun   := FALSE;
            eStateInt  := E_DL_TwoSpeedState.eRunLow;
        END_IF

    E_DL_TwoSpeedState.eFault:
        bOutLowInt  := FALSE;        // 故障相双绕组全断（降级语义已声明 R191）/ Both off, declared
        bOutHighInt := FALSE;
        (* 解除路径（R152 自证可达）：复位沿 AND 双反馈均断 AND 组态已改对 *)
        IF fbTrigReset.Q AND (NOT bFbHigh) AND (NOT bFbLow) AND (NOT bCfgBad) THEN
            bAdhesionInt := FALSE;
            bFbFailInt   := FALSE;
            uErrorId     := 16#0000_0000;
            eStateInt    := E_DL_TwoSpeedState.eIdle;
        END_IF

    ELSE
        (* 非法状态拦截：双断 + 迁兜底态（复用组态段码位） *)
        eStateInt   := E_DL_TwoSpeedState.eFault;
        uErrorId    := 16#0003_050D;
        bErrorInt   := TRUE;
        bOutLowInt  := FALSE;
        bOutHighInt := FALSE;

END_CASE;

(*------------------------------------------------------------------------------
 * 段 6｜反馈校验到期消化：投入命令已发而反馈超时未到 -> 校验失败锁存 + 断该绕组
 *      Feedback verify expiry: command on but feedback never arrived
 *      拍 N 进入：tonFb*.Q 首次为真；本拍行为：锁存 + 断输出 + 迁 eFault；
 *      拍 N+1 转出：eFault 相复位沿 + 双反馈均断解除
 *-----------------------------------------------------------------------------*)
IF tonFbLow.Q AND (eStateInt = E_DL_TwoSpeedState.eRunLow) THEN
    bFbFailInt := TRUE;          // 低速反馈校验失败 / Low feedback verify failed
    uErrorId   := 16#0003_050C;
    bErrorInt  := TRUE;
    bOutLowInt := FALSE;         // 安全侧断该绕组 / Cut the winding on safe side
    eStateInt  := E_DL_TwoSpeedState.eFault;
END_IF

IF tonFbHigh.Q AND (eStateInt = E_DL_TwoSpeedState.eRunHigh) THEN
    bFbFailInt := TRUE;          // 高速反馈校验失败（安全侧断高速）/ High verify failed, cut high
    uErrorId   := 16#0003_050C;
    bErrorInt  := TRUE;
    bOutHighInt := FALSE;
    eStateInt  := E_DL_TwoSpeedState.eFault;
END_IF

(*------------------------------------------------------------------------------
 * 段 7｜输出单一出口（范式 P-05）：两绕组互斥交叉硬闸（结构 + 出口双保险）
 *      Single output exit: cross hard gate, structural plus exit double insurance
 *-----------------------------------------------------------------------------*)
bOutLow  := bOutLowInt AND (NOT bOutHighInt);
bOutHigh := bOutHighInt AND (NOT bOutLowInt);

bSwitching  := (eStateInt = E_DL_TwoSpeedState.eSwUp) OR (eStateInt = E_DL_TwoSpeedState.eSwDown);
bAdhesion   := bAdhesionInt;
bFbFail     := bFbFailInt;
bError      := bErrorInt OR (eStateInt = E_DL_TwoSpeedState.eFault);
eState      := eStateInt;
END_FUNCTION_BLOCK

(* ---- FB_DL_UltrasonicWeldCtrl.st ---- *)
(*
  ==================================================================
  组件名 Component  : FB_DL_UltrasonicWeldCtrl
  分类   Category   : DL_Device
  复杂度 Complexity  : cx5
  版本   Version    : 1.0.0
  功能   Purpose    : 超声波焊接顺控。相位机 eIdle → eDown → eHold → eSonicOn →
                      eCool → eUp → eDone / eFault；能量积分用梯形法（E += (P +
                      Pprev)/2·dt）；超能量 / 欠能量双判据独立成因（R190）+ 超时
                      看门狗；输出 bSonicActive / bWeldDone / fEnergy。
  来源   Source     : t2-2-lbp
  溯源   Origin     : IEC 61131-3 标准语义的道莅防御性实现；超声焊接能量 / 振幅 /
                      时间三模终点为通用工艺语义，clean-room 自研实现，未复制任何
                      闭源代码行。
  平台   Platform   : 纯 IEC 61131-3（TON / R_TRIG / LREAL，无私有库）
  作者   Author     : 道莅代码库 · PLC 编程专家（R56）
  ------------------------------------------------------------------
  同拍多窗说明（R100）：五个窗互斥 —— 每窗 IN 串「本相」闸，任一时刻只有一个窗
                      在计时；配比约束 tSonicTo > tWeld 在组态域闸内判故障
                      （看门狗窗必须覆盖目标窗）。
  边界 Boundary     :
                      一 本件只出焊接命令与能量结算，不驱动换能器电源、不控气缸
                         （属主边界）；
                      二 相级看门狗使能只用相驻留本身（R145）；
                      三 能量梯形积分仅在 eSonicOn 相执行；进入该相时能量清零
                         （单点入口赋值，防跨批残留）；
                      四 故障锁存解除路径 = bReset 上升沿（唯一路径，R188）；
                      五 无全局变量、无外部变量声明、无物理地址寻址。
  输出契约 Output contract:
                      fAmplitudeCmd 恒在 [0, fAmpMax]；fEnergy 为最近一次焊接结算
                      能量 [焦]；bWeldDone 为单拍脉冲（R187 两段式）；
                      eFault 为锁存回放；ePhaseBad 为非法相位兜底专用成员（R128）。
  修订记录 Revision  :
    2026-11-20  v1.0.0  R56 首版（批 4 · 序号 18）
  ==================================================================
*)

TYPE E_DL_UwcPhase :
(
    eIdle    := 0,  // 空闲：等启动沿 / idle, waiting for the start edge
    eDown    := 10, // 下压：等到位反馈 / down, waiting for the position feedback
    eHold    := 20, // 保压：保压计时 / holding, the hold timing
    eSonicOn := 30, // 超声：能量积分与双判据 / sonic on, the energy integral with the twin verdicts
    eCool    := 40, // 冷却：冷却计时 / cooling, the cool timing
    eUp      := 50, // 回升：等原位反馈 / up, waiting for the home feedback
    eDone    := 60, // 完成：结算驻留 / done, the settlement holds
    eFault   := 90  // 故障：成因锁存，超声撤 / fault, the cause is latched with the sonic off
);
END_TYPE

TYPE E_DL_UwcFault :
(
    eNone         := 0, // 无成因 / no cause
    eEnergyHigh   := 1, // 能量超上限（故障级，与 bError 配对）/ the energy is over the ceiling, fault grade paired with bError
    eEnergyLow    := 2, // 焊接窗耗尽能量仍低于下限（故障级，与 bError 配对）/ the window expired with the energy below the floor, fault grade paired with bError
    eSonicTimeout := 3, // 超声相看门狗超时（故障级，与 bError 配对）/ the sonic phase watchdog timed out, fault grade paired with bError
    eDownTimeout  := 4, // 下压相超时（故障级，与 bError 配对）/ the down phase timed out, fault grade paired with bError
    eUpTimeout    := 5, // 回升相超时（故障级，与 bError 配对）/ the up phase timed out, fault grade paired with bError
    eSensorBad    := 6, // 功率非有限或组态非法（故障级，与 bError 配对）/ the power is non finite or the config illegal, fault grade paired with bError
    ePhaseBad     := 7  // 非法相位兜底（故障级，与 bError 配对）/ illegal phase fallback, fault grade paired with bError
);
END_TYPE

FUNCTION_BLOCK FB_DL_UltrasonicWeldCtrl
VAR_INPUT
    bEnable     : BOOL := TRUE;    // 使能，失能时停顺控回空闲 [-] / enable, the sequence stops when disabled
    bReset      : BOOL := FALSE;   // 复位上升沿清故障锁存 [-] / reset rising edge clears the fault latch
    bStart      : BOOL := FALSE;   // 焊接启动脉冲，上升沿受理 [-] / the weld start pulse, accepted on the rising edge
    bAbort      : BOOL := FALSE;   // 中止（电平），任何中间态撤超声回空闲 [-] / the abort level, any middle phase withdraws the sonic
    bPosDownFb  : BOOL := FALSE;   // 焊接位置到位反馈 [-] / the weld position feedback
    bPosUpFb    : BOOL := TRUE;    // 原位反馈 [-] / the home position feedback
    fPowerW     : LREAL := 0.0;    // 超声功率实测 [瓦] / the measured sonic power [watt]
    fAmpSet     : LREAL := 60.0;   // 振幅设定 [百分比]，域 0..100 / the amplitude setpoint [percent], domain zero to one hundred
    fAmpMax     : LREAL := 100.0;  // 振幅上限 [百分比] / the amplitude ceiling [percent]
    fEnergyMinJ : LREAL := 50.0;   // 能量下限 [焦] / the energy floor [joule]
    fEnergyTgtJ : LREAL := 200.0;  // 能量目标 [焦]，域 大于下限 / the energy target [joule], above the floor
    fEnergyMaxJ : LREAL := 300.0;  // 能量上限 [焦]，域 大于目标 / the energy ceiling [joule], above the target
    tHold       : TIME := T#500MS; // 保压时长 [毫秒] / the hold duration [millisecond]
    tWeld       : TIME := T#3S;    // 焊接目标窗 [毫秒] / the weld target window [millisecond]
    tSonicTo    : TIME := T#5S;    // 超声相看门狗窗 [毫秒]，域 大于 tWeld / the sonic watchdog window, above the weld window
    tCool       : TIME := T#1S;    // 冷却时长 [毫秒] / the cool duration [millisecond]
    tDownTo     : TIME := T#5S;    // 下压超时窗 [毫秒] / the down timeout window [millisecond]
    tUpTo       : TIME := T#5S;    // 回升超时窗 [毫秒] / the up timeout window [millisecond]
    fDtS        : LREAL := 0.01;   // 调用周期 [秒]，域 大于零 / the call period [second], domain above zero
END_VAR
VAR_OUTPUT
    bSonicActive  : BOOL := FALSE; // 超声激活命令（相位派生电平）[-] / the sonic active command, a phase derived level
    fAmplitudeCmd : LREAL := 0.0;  // 振幅命令输出 [百分比] / the amplitude command outlet [percent]
    bWeldDone     : BOOL := FALSE; // 焊接完成单拍脉冲 [-] / the weld done single shot pulse
    fEnergy       : LREAL := 0.0;  // 最近一次焊接结算能量 [焦] / the settled energy of the last weld [joule]
    ePhase        : E_DL_UwcPhase := E_DL_UwcPhase.eIdle; // 相位出口 [枚举] / phase outlet [enum]
    eFault        : E_DL_UwcFault := E_DL_UwcFault.eNone; // 成因出口，锁存回放 [枚举] / cause outlet replayed from the latch [enum]
    bError        : BOOL := FALSE; // 故障锁存标志 [-] / fault latch flag
END_VAR
VAR
    rtStart  : R_TRIG; // 启动沿检测，段 0 无条件刷新 / start edge, refreshed unconditionally in segment zero
    rtReset  : R_TRIG; // 复位沿检测，段 0 无条件刷新 / reset edge, refreshed unconditionally in segment zero
    tonDown  : TON;    // 下压超时窗，段 0 无条件刷新 / the down timeout window, refreshed unconditionally
    tonHold  : TON;    // 保压计时窗，段 0 无条件刷新 / the hold timing window, refreshed unconditionally
    tonWeld  : TON;    // 焊接目标窗，段 0 无条件刷新 / the weld target window, refreshed unconditionally
    tonSonic : TON;    // 超声看门狗窗，段 0 无条件刷新 / the sonic watchdog window, refreshed unconditionally
    tonCool  : TON;    // 冷却计时窗，段 0 无条件刷新 / the cool timing window, refreshed unconditionally
    tonUp    : TON;    // 回升超时窗，段 0 无条件刷新 / the up timeout window, refreshed unconditionally
    _ePhase  : E_DL_UwcPhase := E_DL_UwcPhase.eIdle; // 内部相位，CASE 唯一写入目标 / internal phase, the only CASE write target
    _eFaulC  : E_DL_UwcFault := E_DL_UwcFault.eNone; // 故障级成因，锁存至复位沿 / fault cause, latched until the reset edge
    _bFault  : BOOL := FALSE; // 故障锁存位 [-] / fault latch bit
    _bInit   : BOOL := FALSE; // 首扫初始化完成标志（R310）/ first scan initialisation flag
    _bDoneInt: BOOL := FALSE; // 完成脉冲内部位，统一出口映射 / internal done bit, mapped at the unified outlet
    _bInOk   : BOOL := FALSE; // 功率有限 [-] / the power is finite
    _bCfgOk  : BOOL := FALSE; // 组态参数域内 [-] / the configuration is inside the domain
    _fPwPrev : LREAL := 0.0;  // 上拍功率快照 [瓦] / previous scan power snapshot [watt]
    _fEnergyW: LREAL := 0.0;  // 能量积分工作值 [焦] / the energy integral working value [joule]
    _fAmpUse : LREAL := 60.0;  // 钳定后的振幅 [百分比] / the clamped amplitude [percent]
END_VAR

// 段 0｜定时器与沿检测无条件周期刷新（禁入分支），IN 只串相位闸与故障闸（FB50-1）/ segment 0, unconditional refresh, no instance call inside a branch
rtStart(CLK := bStart); // 启动沿 / the start edge
rtReset(CLK := bReset); // 复位沿 / the reset edge
tonDown(IN := (_ePhase = E_DL_UwcPhase.eDown) AND (NOT _bFault), PT := tDownTo); // 下压超时窗 / the down timeout window
tonHold(IN := (_ePhase = E_DL_UwcPhase.eHold) AND (NOT _bFault), PT := tHold); // 保压计时窗 / the hold timing window
tonWeld(IN := (_ePhase = E_DL_UwcPhase.eSonicOn) AND (NOT _bFault), PT := tWeld); // 焊接目标窗 / the weld target window
tonSonic(IN := (_ePhase = E_DL_UwcPhase.eSonicOn) AND (NOT _bFault), PT := tSonicTo); // 超声看门狗窗 / the sonic watchdog window
tonCool(IN := (_ePhase = E_DL_UwcPhase.eCool) AND (NOT _bFault), PT := tCool); // 冷却计时窗 / the cool timing window
tonUp(IN := (_ePhase = E_DL_UwcPhase.eUp) AND (NOT _bFault), PT := tUpTo); // 回升超时窗 / the up timeout window

// 段 1｜首扫初始化（R310）/ segment 1, first scan initialisation
IF NOT _bInit THEN // 首扫一拍 / the very first scan
    _bInit := TRUE; // 置首扫完成标志 / raise the first scan flag
    _ePhase := E_DL_UwcPhase.eIdle; // 相位从空闲起步 / the phase starts from idle
    _eFaulC := E_DL_UwcFault.eNone; // 故障级成因清零 / clear the fault cause
    _bFault := FALSE; // 故障锁存清零 / clear the fault latch
    _fPwPrev := fPowerW; // 快照取当拍 / the snapshot takes this scan
END_IF

// 段 2｜复位沿作用域：清锁存 / 迁相位 / 清能量工作值（三项逐项声明）/ segment 2, reset edge scope declared item by item
IF rtReset.Q THEN // 复位沿 / the reset edge
    _bFault := FALSE; // 作用域一：清故障锁存 / scope one, clear the fault latch
    _eFaulC := E_DL_UwcFault.eNone; // 作用域一：清故障级成因 / scope one, clear the fault cause
    _ePhase := E_DL_UwcPhase.eIdle; // 作用域二：迁回空闲相 / scope two, migrate back to idle
    _fEnergyW := 0.0; // 作用域三：清能量工作值（结算出口 fEnergy 保持）/ scope three, the integral clears while the settlement holds
END_IF

// 段 3｜组态与输入域闸（R151 全覆盖，含 R100 配比）/ segment 3, the configuration gate with the window pairing
_bInOk := (fPowerW = fPowerW) AND ((fPowerW - fPowerW) = (fPowerW - fPowerW)) AND (fPowerW >= 0.0); // 功率有限且非负 / the power is finite and non negative
_bCfgOk := (fAmpSet >= 0.0) AND (fAmpSet = fAmpSet) AND (fAmpMax > 0.0) AND (fAmpMax = fAmpMax) AND (fEnergyMinJ > 0.0) AND (fEnergyMinJ = fEnergyMinJ) AND (fEnergyTgtJ > fEnergyMinJ) AND (fEnergyTgtJ = fEnergyTgtJ) AND (fEnergyMaxJ > fEnergyTgtJ) AND (fEnergyMaxJ = fEnergyMaxJ) AND (tHold > T#0S) AND (tWeld > T#0S) AND (tSonicTo > tWeld) AND (tCool > T#0S) AND (tDownTo > T#0S) AND (tUpTo > T#0S) AND (fDtS > 0.0) AND (fDtS = fDtS); // 组态参数域判定（含 tSonicTo > tWeld 配比，R100）/ the configuration verdict with the pairing
IF (NOT _bInOk) OR (NOT _bCfgOk) THEN // 功率无效或组态非法 / a void power or an illegal configuration
    IF NOT _bFault THEN // 未锁存才迁移（防同拍抹除）/ migrate only while unlatched
        _bFault := TRUE; // 置故障锁存 / raise the fault latch
        _eFaulC := E_DL_UwcFault.eSensorBad; // 故障级成因（R45 配对 bError）/ the fault cause paired with bError
        _ePhase := E_DL_UwcPhase.eFault; // 迁故障相 / migrate to the fault phase
    END_IF
END_IF
_fAmpUse := fAmpSet; // 振幅直通 / the amplitude passes through
IF _fAmpUse > fAmpMax THEN // 振幅上钳（R117 两级回退）/ clamp the amplitude high
    _fAmpUse := fAmpMax; // 钳到上限 / clamp to the ceiling
END_IF

// 段 4｜相位机：ENUM + CASE，含 ELSE 非法相位兜底（R128）/ segment 4, the phase machine with an ELSE fallback
CASE _ePhase OF
E_DL_UwcPhase.eIdle: // 空闲相：等启动沿 / the idle phase, waiting for the start edge
    IF bEnable AND (NOT _bFault) AND (NOT bAbort) AND rtStart.Q THEN // 启动沿受理 / the start edge is accepted
        _fEnergyW := 0.0; // 能量工作值清零 / clear the energy integral
        _fPwPrev := 0.0; // 功率快照清零 / clear the power snapshot
        _ePhase := E_DL_UwcPhase.eDown; // 迁下压相 / migrate to the down phase
    END_IF

E_DL_UwcPhase.eDown: // 下压相：等到位反馈（退出条件 ≥2：到位 / 超时 / 中止 / 失能，R98）/ the down phase with at least two exit conditions
    IF (NOT bEnable) OR bAbort THEN // 失能或中止 / disabled or aborting
        _ePhase := E_DL_UwcPhase.eIdle; // 回空闲相 / back to idle
    ELSIF bPosDownFb THEN // 到位 / the position is reached
        _ePhase := E_DL_UwcPhase.eHold; // 迁保压相 / migrate to the hold phase
    ELSIF tonDown.Q THEN // 下压超时 / the down phase timed out
        _bFault := TRUE; // 置故障锁存 / raise the fault latch
        _eFaulC := E_DL_UwcFault.eDownTimeout; // 故障级成因（R45 配对 bError）/ the fault cause paired with bError
        _ePhase := E_DL_UwcPhase.eFault; // 迁故障相 / migrate to the fault phase
    END_IF

E_DL_UwcPhase.eHold: // 保压相：保压计时 / the hold phase, the hold timing
    IF (NOT bEnable) OR bAbort THEN // 失能或中止 / disabled or aborting
        _ePhase := E_DL_UwcPhase.eIdle; // 回空闲相 / back to idle
    ELSIF tonHold.Q THEN // 保压时长已到 / the hold duration elapsed
        _fEnergyW := 0.0; // 能量积分入口清零（单点入口赋值，防跨批残留）/ the entry zeroing of the energy integral
        _fPwPrev := 0.0; // 功率快照入口清零 / the entry zeroing of the power snapshot
        _ePhase := E_DL_UwcPhase.eSonicOn; // 迁超声相 / migrate to the sonic phase
    END_IF

E_DL_UwcPhase.eSonicOn: // 超声相：梯形能量积分 + 双判据 + 看门狗 / the sonic phase, the trapezoid integral with the twin verdicts and the watchdog
    IF (NOT bEnable) OR bAbort THEN // 失能或中止 / disabled or aborting
        _ePhase := E_DL_UwcPhase.eIdle; // 回空闲相 / back to idle
    ELSE // 焊接中 / welding
        IF _bInOk THEN // 功率有限 / the power is finite
            _fEnergyW := _fEnergyW + (fPowerW + _fPwPrev) / 2.0 * fDtS; // 梯形法能量积分，除子无（乘法口径）/ the trapezoid energy integral
            _fPwPrev := fPowerW; // 功率快照推进 / advance the power snapshot
        END_IF
        fEnergy := _fEnergyW; // 能量出口实时跟随 / the energy outlet follows live
        IF _fEnergyW > fEnergyMaxJ THEN // 超能量判据（R190 独立成因）/ the over energy criterion, an independent cause
            _bFault := TRUE; // 置故障锁存 / raise the fault latch
            _eFaulC := E_DL_UwcFault.eEnergyHigh; // 故障级成因（R45 配对 bError）/ the fault cause paired with bError
            _ePhase := E_DL_UwcPhase.eFault; // 迁故障相 / migrate to the fault phase
        ELSIF tonSonic.Q THEN // 看门狗超时（覆盖目标窗的兜底，R100）/ the watchdog expired, the fallback over the target window
            _bFault := TRUE; // 置故障锁存 / raise the fault latch
            _eFaulC := E_DL_UwcFault.eSonicTimeout; // 故障级成因（R45 配对 bError）/ the fault cause paired with bError
            _ePhase := E_DL_UwcPhase.eFault; // 迁故障相 / migrate to the fault phase
        ELSIF tonWeld.Q THEN // 焊接目标窗耗尽 / the weld target window expired
            IF _fEnergyW < fEnergyMinJ THEN // 欠能量判据（R190 独立成因）/ the under energy criterion, an independent cause
                _bFault := TRUE; // 置故障锁存 / raise the fault latch
                _eFaulC := E_DL_UwcFault.eEnergyLow; // 故障级成因（R45 配对 bError）/ the fault cause paired with bError
                _ePhase := E_DL_UwcPhase.eFault; // 迁故障相 / migrate to the fault phase
            ELSE // 能量在窗内，按时间终点收焊 / the energy is inside the window, the time based close
                _ePhase := E_DL_UwcPhase.eCool; // 迁冷却相 / migrate to the cool phase
            END_IF
        ELSIF _fEnergyW >= fEnergyTgtJ THEN // 能量达标（优先终点）/ the energy target is reached, the primary end
            _ePhase := E_DL_UwcPhase.eCool; // 迁冷却相 / migrate to the cool phase
        END_IF
    END_IF

E_DL_UwcPhase.eCool: // 冷却相：冷却计时 / the cool phase, the cool timing
    IF (NOT bEnable) OR bAbort THEN // 失能或中止 / disabled or aborting
        _ePhase := E_DL_UwcPhase.eIdle; // 回空闲相 / back to idle
    ELSIF tonCool.Q THEN // 冷却时长已到 / the cool duration elapsed
        _ePhase := E_DL_UwcPhase.eUp; // 迁回升相 / migrate to the up phase
    END_IF

E_DL_UwcPhase.eUp: // 回升相：等原位反馈（退出条件 ≥2：原位 / 超时 / 中止 / 失能，R98）/ the up phase with at least two exit conditions
    IF (NOT bEnable) OR bAbort THEN // 失能或中止 / disabled or aborting
        _ePhase := E_DL_UwcPhase.eIdle; // 回空闲相 / back to idle
    ELSIF bPosUpFb THEN // 原位 / the home position is reached
        _bDoneInt := TRUE; // 完成脉冲内部位置位（统一出口映射，R187）/ raise the internal done bit
        _ePhase := E_DL_UwcPhase.eDone; // 迁完成相 / migrate to the done phase
    ELSIF tonUp.Q THEN // 回升超时 / the up phase timed out
        _bFault := TRUE; // 置故障锁存 / raise the fault latch
        _eFaulC := E_DL_UwcFault.eUpTimeout; // 故障级成因（R45 配对 bError）/ the fault cause paired with bError
        _ePhase := E_DL_UwcPhase.eFault; // 迁故障相 / migrate to the fault phase
    END_IF

E_DL_UwcPhase.eDone: // 完成相：结算驻留，等复位或新启动 / the done phase, the settlement holds until reset or a new start
    IF (NOT bEnable) OR rtStart.Q THEN // 失能或新启动沿 / disabled or a new start edge
        _ePhase := E_DL_UwcPhase.eIdle; // 回空闲相 / back to idle
    END_IF

E_DL_UwcPhase.eFault: // 故障相：超声撤，成因锁存，等复位沿 / the fault phase, the sonic off until the reset edge
    IF NOT bEnable THEN // 失能 / disabled
        _ePhase := E_DL_UwcPhase.eIdle; // 迁未使能相 / migrate to idle
    END_IF

ELSE // 非法相位兜底（R128）/ the illegal phase fallback
    _bFault := TRUE; // 置故障锁存 / raise the fault latch
    _eFaulC := E_DL_UwcFault.ePhaseBad; // 故障级成因（R45 配对 bError）/ the fault cause paired with bError
    _ePhase := E_DL_UwcPhase.eFault; // 迁故障相 / migrate to the fault phase
END_CASE

// 段 6｜命令出口派生（互斥的结构性承载）/ segment 6, the command outlets, the structural carrier
bSonicActive := (_ePhase = E_DL_UwcPhase.eSonicOn) AND (NOT _bFault) AND bEnable AND (NOT bAbort); // 超声激活命令：仅超声相派生 / the sonic command, derived in the sonic phase only
IF bSonicActive THEN // 超声激活拍 / the sonic active scan
    fAmplitudeCmd := _fAmpUse; // 振幅命令出口 / the amplitude command outlet
ELSE // 非激活拍 / the inactive scan
    fAmplitudeCmd := 0.0; // 振幅归零（安全侧）/ the amplitude zeroes, the safe side
END_IF

// 段 7｜统一出口 / segment 7, the unified outlet
bWeldDone := _bDoneInt; // 完成脉冲映射本拍值 / map the done pulse for this scan
_bDoneInt := FALSE; // 映射后立即撤销，保证单拍宽度（R187 两段式）/ revoke right after mapping
IF _bFault THEN // 故障锁存优先 / the fault latch takes priority
    eFault := _eFaulC; // 故障级成因锁存回放（R152）/ the fault cause replayed from the latch
ELSE
    eFault := E_DL_UwcFault.eNone; // 无锁存即无成因 / no latch, no cause
END_IF
ePhase := _ePhase; // 相位出口单点映射 / single point phase outlet mapping
bError := _bFault; // 故障标志与锁存位同源 / the fault flag shares the latch source
END_FUNCTION_BLOCK

(* ---- FB_DL_UncoilerMandrelSeq.st ---- *)
(*
  Name: FB_DL_UncoilerMandrelSeq
  Category: DL_Device
  Version: 1.0.0
  Round: R89 / 2026-11-25
  开源溯源：clean-room 自研（族 板带剪切分条卷取，ST 开源生态实测 0 命中，无外部代码引入）
  功能：开卷机卷筒胀缩与压辊顺序：压辊压下→卷筒胀径→对中确认→允许穿带。
  边界条件：① 卷径与设定值过非有限闸；越域即故障（101）；
            ② 压辊/胀径/对中三相各用独立 TON，PT 均取 tTimeoutS，禁跨相共用（R100）；
            ③ 胀径确认用差值容差比较（±0.5 mm），禁浮点判等；
            ④ 故障解除唯一路径：故障相内 xStart 释放（R152），清锁存回 eIdle。
  状态机：eIdle / ePressRoll / eExpand / eCenter / eReady / eFault（CASE 含 ELSE 兜底）。
*)
TYPE E_DL_UmsPhase :
(
    eIdle      := 0,    (* 待机：等启动沿 / Idle, waiting for start edge *)
    ePressRoll := 10,   (* 压辊相：等压下反馈 / Press roll, waiting down feedback *)
    eExpand    := 20,   (* 胀径相：等卷筒胀到设定 / Expanding to diameter setpoint *)
    eCenter    := 30,   (* 对中相：等对中确认 / Centering confirmation *)
    eReady     := 40,   (* 就绪相：允许穿带 / Ready, strip threading allowed *)
    eFault     := 90    (* 故障相：锁存待释放 / Fault latched, awaiting release *)
);
END_TYPE

FUNCTION_BLOCK FB_DL_UncoilerMandrelSeq
VAR_INPUT
    xStart : BOOL;              (* 启动命令（上升沿起序） [-] Start command, rising edge *)
    fMandrelDiaMm : REAL;       (* 卷筒胀径实测 [mm] Mandrel diameter actual [mm] *)
    fMandrelDiaSetMm : REAL;    (* 卷筒胀径设定 [mm] Mandrel diameter setpoint [mm] *)
    xPressRollDown : BOOL;      (* 压辊压下到位反馈 [-] Press roll down feedback *)
    xCentered : BOOL;           (* 对中确认反馈 [-] Centering feedback *)
    tTimeoutS : TIME;           (* 单相超时窗 [ms] Phase timeout window [ms] *)
END_VAR
VAR_OUTPUT
    eState : E_DL_UmsPhase;     (* 当前相 [-] Present phase *)
    xReady : BOOL;              (* 允许穿带 [-] Ready for strip threading *)
    xFault : BOOL;              (* 故障锁存标志 [-] Fault latched *)
    nErrCode : INT;             (* 故障码 0/101 组态/102~104 超时/105 非法相 [-] Error code *)
END_VAR
VAR
    _ePhase : E_DL_UmsPhase := E_DL_UmsPhase.eIdle;  (* 内部相（CASE 唯一写入目标） [-] Internal phase *)
    _bFaultLatch : BOOL := FALSE;   (* 故障锁存位 [-] Fault latch *)
    _bReqFault : BOOL := FALSE;     (* 单拍故障请求（段 1 预清） [-] Fault request *)
    _bCfgBad : BOOL := FALSE;       (* 组态非法当拍量 [-] Configuration bad *)
    _nErr : INT := 0;               (* 故障码锁存 [-] Latched error code *)
    _nReqErr : INT := 0;            (* 当拍请求码 [-] Requested error code *)
    _fDiaErrMm : REAL := 0.0;       (* 胀径偏差绝对量 [mm] Absolute diameter deviation [mm] *)
    tonPress : TON;                 (* 压辊超时（段 0 无条件调用） / Press roll timeout *)
    tonExpand : TON;                (* 胀径超时（段 0 无条件调用） / Expand timeout *)
    tonCenter : TON;                (* 对中超时（段 0 无条件调用） / Centering timeout *)
    rtStart : R_TRIG;               (* 启动沿（段 0 无条件调用） / Start edge *)
END_VAR
VAR CONSTANT
    DL_UMS_TOL : REAL := 0.5;       (* 胀径到位容差 [mm] Diameter tolerance [mm] *)
END_VAR
(* —— 段 0：沿与三 TON 无条件周期刷新（R7），IN 仅由相位派生 —— *)
rtStart(CLK := xStart);                                                     (* 启动沿 / Start edge *)
tonPress(IN := (_ePhase = E_DL_UmsPhase.ePressRoll), PT := tTimeoutS);      (* 压辊超时 / Press timeout *)
tonExpand(IN := (_ePhase = E_DL_UmsPhase.eExpand), PT := tTimeoutS);        (* 胀径超时 / Expand timeout *)
tonCenter(IN := (_ePhase = E_DL_UmsPhase.eCenter), PT := tTimeoutS);        (* 对中超时 / Centering timeout *)
(* 非有限闸（NaN 自反 + Inf 差值自减）+ 组态域闸：两浮点入参全枚举（R272） *)
_bCfgBad := (fMandrelDiaMm <> fMandrelDiaMm) OR ((fMandrelDiaMm - fMandrelDiaMm) <> 0.0)
         OR (fMandrelDiaSetMm <> fMandrelDiaSetMm) OR ((fMandrelDiaSetMm - fMandrelDiaSetMm) <> 0.0)
         OR (fMandrelDiaSetMm < 300.0) OR (fMandrelDiaSetMm > 2200.0)
         OR (fMandrelDiaMm < 100.0) OR (fMandrelDiaMm > 2300.0) OR (tTimeoutS <= T#0S);
(* 胀径偏差绝对量：容差比较用差值，禁浮点判等 *)
_fDiaErrMm := ABS(fMandrelDiaMm - fMandrelDiaSetMm);
(* —— 段 1：单拍量预清零 —— *)
_bReqFault := FALSE;
_nReqErr := 0;
IF _bCfgBad THEN
    _bReqFault := TRUE; _nReqErr := 101;        (* 组态非法 / Configuration bad *)
END_IF
(* —— 段 2：故障锁存解除（唯一路径 = 故障相内 xStart 释放，R152） —— *)
IF _bFaultLatch AND (NOT xStart) THEN
    _bFaultLatch := FALSE;                      (* 清锁存 / Clear latch *)
    _nErr := 0;                                 (* 清码 / Clear code *)
    _ePhase := E_DL_UmsPhase.eIdle;             (* 迁回待机 / Back to idle *)
END_IF
(* —— 段 3：主状态机（ENUM + CASE，ELSE 兜底） —— *)
CASE _ePhase OF
E_DL_UmsPhase.eIdle:
    IF rtStart.Q AND (NOT _bFaultLatch) THEN
        _ePhase := E_DL_UmsPhase.ePressRoll;    (* 起序 → 压辊压下 / Start, press roll down *)
    END_IF
E_DL_UmsPhase.ePressRoll:
    IF xPressRollDown THEN
        _ePhase := E_DL_UmsPhase.eExpand;       (* 压辊到位 → 胀径 / Pressed, expand *)
    ELSIF tonPress.Q THEN
        _bReqFault := TRUE; _nReqErr := 102;    (* 压辊超时 / Press roll timeout *)
    END_IF
E_DL_UmsPhase.eExpand:
    IF _fDiaErrMm <= DL_UMS_TOL THEN
        _ePhase := E_DL_UmsPhase.eCenter;       (* 胀到设定 → 对中 / Expanded, center *)
    ELSIF tonExpand.Q THEN
        _bReqFault := TRUE; _nReqErr := 103;    (* 胀径超时 / Expand timeout *)
    END_IF
E_DL_UmsPhase.eCenter:
    IF xCentered THEN
        _ePhase := E_DL_UmsPhase.eReady;        (* 对中确认 → 就绪 / Centered, ready *)
    ELSIF tonCenter.Q THEN
        _bReqFault := TRUE; _nReqErr := 104;    (* 对中超时 / Centering timeout *)
    END_IF
E_DL_UmsPhase.eReady:
    IF NOT xStart THEN
        _ePhase := E_DL_UmsPhase.eIdle;         (* 启动释放 → 待机（撤穿带许可） / Start released *)
    END_IF
E_DL_UmsPhase.eFault:
    _fDiaErrMm := ABS(fMandrelDiaMm - fMandrelDiaSetMm);   (* 故障相驻留：仅刷新偏差量供追溯 *)
ELSE
    _bReqFault := TRUE;                         (* 非法相兜底 / Illegal phase fallback *)
    _nReqErr := 105;
END_CASE
(* —— 段 4：故障请求统一落地（唯一锁存点 + 同步迁相，R187/R252） —— *)
IF _bReqFault AND (NOT _bFaultLatch) THEN
    _bFaultLatch := TRUE;                       (* 锁存 / Latch *)
    _nErr := _nReqErr;                          (* 码锁存回放 / Latched code *)
    _ePhase := E_DL_UmsPhase.eFault;            (* 同步迁相 / Migrate to fault *)
END_IF
(* —— 段 5：统一出口（各出口单点赋值） —— *)
eState := _ePhase;
xReady := (_ePhase = E_DL_UmsPhase.eReady) AND (NOT _bFaultLatch);
xFault := _bFaultLatch;
nErrCode := _nErr;
END_FUNCTION_BLOCK

(* ---- FB_DL_UnlockHoldTimeout.st ---- *)
(*
  Component : FB_DL_UnlockHoldTimeout
  Category  : DL_Device
  Type      : FB
  Version   : 1.0.0
  CodeSeg   : 16#03_1_02
  Summary   : 安全门解锁保持超时监视：解锁有效但门未开持续超阈 → 电磁铁/机械卡滞提示，事件沿计数留痕。
              Door unlock hold timeout monitor: unlocked but not opened over limit, solenoid or jam hint with edge-counted ledger.
  溯源声明  : 道莅自研 clean-room
  边界安全  : 只消费 FB_DL_GuardLockDoor 对外输出引脚（不侵入其内部状态）；超时阈值 tHoldLimMs
              提为输入引脚（带 ms 单位，禁魔法数）并做正域闸（> 0，防 TON 无效整定）；
              提示为非锁存自清（条件消失即清），事件计数走上升沿防电平重复累加；
              TON 每拍无条件刷新（段 0）；全浮点比较带 fEps 容差。
  复用      : 消费 FB_DL_GuardLockDoor 的对外输出引脚（bUnlockActive / bDoorOpened），无实例依赖
*)

FUNCTION_BLOCK FB_DL_UnlockHoldTimeout
VAR_INPUT
    bRun          : BOOL;              (* 监视使能 · Enable *)
    bUnlockActive : BOOL;              (* 解锁有效输出 [开关]，来自门控 FB 对外引脚 · Unlock active from door FB *)
    bDoorOpened   : BOOL;              (* 门已开开关 [开关] · Door opened switch *)
    tHoldLimMs    : TIME  := T#3000MS; (* 解锁保持超时阈 [ms] · Hold timeout limit *)
    fEps          : LREAL := 1.0E-6;   (* 浮点判零容差 [实数域] · Floating zero tolerance *)
END_VAR
VAR_OUTPUT
    bHoldNow  : BOOL;                   (* 当前处于超时判据窗口内 [开关] · In the hold judgement window *)
    bJamWarn  : BOOL;                   (* 卡滞提示 [提示]，非锁存自清 · Jam hint, self-clearing *)
    nJamCount : UDINT;                  (* 卡滞事件累计 [次]，沿计数防回卷 · Jam event count *)
    bError    : BOOL;                   (* 故障标志，与故障码配对 · Fault flag paired with codes *)
    uErrorId  : UDINT;                  (* 事件码 16#0000_0102，0 无事件 · Event code *)
END_VAR
VAR
    uCode   : WORD;    (* 码位暂存，每拍重算 [码] · Code staging *)
    tonHold : TON;     (* 解锁保持计时 [ms]，每拍无条件刷新 · Hold timing timer *)
    bWarnPrv: BOOL;    (* 上拍提示快照，事件沿判据 · Previous warn snapshot *)
    nCycles : UDINT;   (* 监视拍计数 [拍]，防回卷 · Monitor scan count *)
END_VAR
VAR CONSTANT
    DL_UHT_WRAP : UDINT := 4294967290;  (* 计数防回卷余量 [次] · Counter wrap guard *)
END_VAR

(* === 段 0 · 实例刷新（每拍无条件，红线 7）=== *)
tonHold(IN := bRun AND bUnlockActive AND (NOT bDoorOpened), PT := tHoldLimMs);
                                        (* 解锁有效且门未开：保持计时 / Hold timing while unlocked and closed *)
bHoldNow := tonHold.Q;                  (* 判据窗口在报状态 / Window active status *)

(* === 段 1 · 输入校验与量程闸 === *)
uCode := 16#0000;                       // 每拍清码（可达清零基线）/ Clear codes each scan
IF tHoldLimMs <= T#0MS THEN
    uCode := 16#0102;                   // 故障级：超时阈非正域，监视失效 / Fault: non-positive limit
END_IF

(* === 段 2 · 主逻辑：保持超时判据（非锁存自清）=== *)
IF bRun AND (uCode = 16#0000) THEN
    bJamWarn := tonHold.Q;              (* 超时到点即提示；解锁或开门条件消失下拍自清 / Hint while timed out *)
    IF bJamWarn AND (NOT bWarnPrv) THEN
        IF nJamCount < DL_UHT_WRAP THEN
            nJamCount := nJamCount + 1; (* 事件上升沿计数，防电平重复累加 / Edge-counted event *)
        END_IF
    END_IF
    IF nCycles < DL_UHT_WRAP THEN
        nCycles := nCycles + 1;         (* 监视拍计数 / Monitor scan count *)
    END_IF
ELSE
    bJamWarn := FALSE;                  (* 撤使能提示清零（可达清零路径）/ Clear on disable *)
END_IF
bWarnPrv := bJamWarn;                   (* 提示快照 / Warn snapshot *)

(* === 段 3 · 输出映射与故障码 === *)
bError := (uCode <> 16#0000) OR bJamWarn;   (* 故障标志：域外码或卡滞提示 / Fault flag *)
IF bJamWarn THEN
    uErrorId := WORD_TO_UDINT(16#0102); (* 码位 16#0000_0102 解锁保持超时 / Hold timeout code *)
ELSE
    uErrorId := WORD_TO_UDINT(uCode);   (* 域外码或零 / Domain code or zero *)
END_IF
END_FUNCTION_BLOCK

(* ---- FB_DL_VacIonizerBalance.st ---- *)
(*
  ==================================================================
  组件名 Component  : FB_DL_VacIonizerBalance
  分类   Category   : DL_Device
  复杂度 Complexity  : cx3
  版本   Version    : 1.0.0
  功能   Purpose    : 离子风机正负离子平衡监视。平衡偏差 = (iP - iN)/( |iP| + |iN| )
                      × 100；正偏 / 负偏双判据独立成因（R190）带迟滞防抖；衰减
                      时间估计：检测到步进突变（|iP| 突变 > fStepThresh）起计时，
                      偏差回带内锁存历时（由采样周期累加），时限 tDecayMax 由
                      TON 判 eDecaySlow；传感器非有限或双低电流判 eSensorBad。
  来源   Source     : t2-2-lbp（ESD 设备族）
  溯源   Origin     : IEC 61131-3 标准语义的道莅防御性实现；离子平衡度与衰减时间
                      为 ESD 公开评价语义（IEC 61340 概念域），clean-room 自研实现，
                      未复制任何闭源代码行。
  平台   Platform   : 纯 IEC 61131-3（TON / R_TRIG / LREAL 运算，无私有库）
  作者   Author     : 道莅代码库 · PLC 编程专家（R56）
  ------------------------------------------------------------------
  边界 Boundary     :
                      一 本件只做平衡判级与衰减估计，不调风机风量、不做高压控制
                         （属主边界）；
                      二 判据方向性（R146）：正偏与负偏为同量纲双向异常，成因独立；
                      三 fDecayS 由采样周期累加估计（秒）；eDecaySlow 由 TON
                         （PT = tDecayMax）判定，两口径职责分离并在头注释声明；
                      四 成因锁存解除路径 = bReset 上升沿（唯一路径，头注释声明，R188）；
                      五 无全局变量、无外部变量声明、无物理地址寻址。
  输出契约 Output contract:
                      fBalDevPct 为平衡偏差百分比；bBalanced 迟滞输出；
                      eFault 为锁存回放；ePhaseBad 为非法相位兜底专用成员（R128）。
  修订记录 Revision  :
    2026-11-20  v1.0.0  R56 首版（批 3 · 序号 11）
  ==================================================================
*)

TYPE E_DL_VibPhase :
(
    eIdle  := 0,  // 未使能：监视停摆 / disabled, the watch is idle
    eRun   := 10, // 运行：逐拍判级 / running, graded every scan
    eDecay := 20, // 衰减测试：步进突变后计时中 / decay test, timing after a step
    eFault := 90  // 故障：成因锁存 / fault, the cause is latched
);
END_TYPE

TYPE E_DL_VibFault :
(
    eNone      := 0, // 无成因 / no cause
    ePosSkew   := 1, // 正偏超限（故障级，与 bError 配对）/ the positive skew is over the limit, fault grade paired with bError
    eNegSkew   := 2, // 负偏超限（故障级，与 bError 配对）/ the negative skew is over the limit, fault grade paired with bError
    eDecaySlow := 3, // 衰减超时（故障级，与 bError 配对）/ the decay outlasted the window, fault grade paired with bError
    eSensorBad := 4, // 传感器非有限或双低电流（故障级，与 bError 配对）/ a sensor is non finite or both currents are void, fault grade paired with bError
    ePhaseBad  := 5  // 非法相位兜底（故障级，与 bError 配对）/ illegal phase fallback, fault grade paired with bError
);
END_TYPE

FUNCTION_BLOCK FB_DL_VacIonizerBalance
VAR_INPUT
    bEnable     : BOOL := TRUE;    // 使能，失能时监视停摆 [-] / enable, the watch stops when disabled
    bReset      : BOOL := FALSE;   // 复位上升沿清全部成因锁存 [-] / reset rising edge clears every cause latch
    iP          : LREAL := 10.0;   // 正离子电流采样 [微安] / the positive ion current sample [microampere]
    iN          : LREAL := 10.0;   // 负离子电流采样 [微安] / the negative ion current sample [microampere]
    fBalLim     : LREAL := 10.0;   // 平衡限（偏差百分比带宽）[百分比]，域 大于零 / the balance limit band [percent], domain above zero
    fHystPct    : LREAL := 2.0;    // 迟滞带宽 [百分比]，域 0..平衡限 / the hysteresis band [percent], inside the limit
    fStepThresh : LREAL := 5.0;    // 衰减测试步进突变阈值 [微安] / the decay test step threshold [microampere]
    tDecayMax   : TIME := T#10S;   // 衰减时限 [毫秒]，域 大于零 / the decay time limit [millisecond], domain above zero
    fDtS        : LREAL := 0.1;    // 调用周期 [秒]，域 大于零 / the call period [second], domain above zero
END_VAR
VAR_OUTPUT
    fBalDevPct : LREAL := 0.0;  // 平衡偏差百分比 [百分比] / the balance deviation [percent]
    bBalanced  : BOOL := FALSE; // 平衡在带内（迟滞输出）[-] / the balance is inside the band, a hysteresis outlet
    fDecayS    : LREAL := 0.0;  // 最近一次衰减历时估计 [秒] / the last decay duration estimate [second]
    ePhase     : E_DL_VibPhase := E_DL_VibPhase.eIdle; // 相位出口 [枚举] / phase outlet [enum]
    eFault     : E_DL_VibFault := E_DL_VibFault.eNone; // 成因出口，锁存回放 [枚举] / cause outlet replayed from the latch [enum]
    bError     : BOOL := FALSE; // 故障锁存标志 [-] / fault latch flag
END_VAR
VAR
    rtReset  : R_TRIG; // 复位沿检测，段 0 无条件刷新 / reset edge, refreshed unconditionally in segment zero
    tonDecay : TON;    // 衰减时限计时，段 0 无条件刷新 / decay limit timer, refreshed unconditionally in segment zero
    _ePhase  : E_DL_VibPhase := E_DL_VibPhase.eIdle; // 内部相位，CASE 唯一写入目标 / internal phase, the only CASE write target
    _eFaulC  : E_DL_VibFault := E_DL_VibFault.eNone; // 故障级成因，锁存至复位沿 / fault cause, latched until the reset edge
    _bFault  : BOOL := FALSE; // 故障锁存位 [-] / fault latch bit
    _bInit   : BOOL := FALSE; // 首扫初始化完成标志（R310）/ first scan initialisation flag
    _bInOk   : BOOL := FALSE; // 两电流输入均有限 [-] / both current inputs are finite
    _bCfgOk  : BOOL := FALSE; // 组态参数域内 [-] / the configuration is inside the domain
    _bBad    : BOOL := FALSE; // 传感器无效锁存 [-] / the sensor bad latch
    _fDen    : LREAL := 0.0;  // 电流幅值和（除子）[微安] / the sum of current magnitudes, the divisor
    _fDev    : LREAL := 0.0;  // 平衡偏差工作值 [百分比] / the balance deviation working value [percent]
    _fIPrev  : LREAL := 0.0;  // 上拍正离子电流快照 [微安] / previous scan positive current snapshot [microampere]
    _fElapS  : LREAL := 0.0;  // 衰减历时累加 [秒] / the decay duration accumulator [second]
    _bPosL   : BOOL := FALSE; // 正偏迟滞锁存 [-] / the positive skew hysteresis latch
    _bNegL   : BOOL := FALSE; // 负偏迟滞锁存 [-] / the negative skew hysteresis latch
END_VAR

// 段 0｜定时器与沿检测无条件周期刷新（禁入分支），IN 只串相位闸与故障闸 / segment 0, unconditional refresh with the phase and fault gates on IN only
rtReset(CLK := bReset); // 复位沿无条件刷新 / unconditional refresh of the reset edge
tonDecay(IN := (_ePhase = E_DL_VibPhase.eDecay) AND (NOT _bFault), PT := tDecayMax); // 衰减时限，IN 串衰减相闸与故障闸 / the decay limit with the phase and fault gates on IN

// 段 1｜首扫初始化（R310）/ segment 1, first scan initialisation
IF NOT _bInit THEN // 首扫一拍 / the very first scan
    _bInit := TRUE; // 置首扫完成标志 / raise the first scan flag
    _ePhase := E_DL_VibPhase.eRun; // 相位从运行起步 / the phase starts in run
    _eFaulC := E_DL_VibFault.eNone; // 故障级成因清零 / clear the fault cause
    _bFault := FALSE; // 故障锁存清零 / clear the fault latch
    _fIPrev := iP; // 快照取当拍 / the snapshot takes this scan
END_IF

// 段 2｜复位沿作用域：清锁存 / 迁相位 / 清迟滞与历时（三项逐项声明）/ segment 2, reset edge scope declared item by item
IF rtReset.Q THEN // 复位沿 / the reset edge
    _bFault := FALSE; // 作用域一：清故障锁存 / scope one, clear the fault latch
    _eFaulC := E_DL_VibFault.eNone; // 作用域一：清故障级成因 / scope one, clear the fault cause
    _bPosL := FALSE; // 作用域一：清正偏迟滞 / scope one, clear the positive latch
    _bNegL := FALSE; // 作用域一：清负偏迟滞 / scope one, clear the negative latch
    _bBad := FALSE; // 作用域一：清传感器无效锁存 / scope one, clear the sensor bad latch
    _ePhase := E_DL_VibPhase.eRun; // 作用域二：迁回运行相 / scope two, migrate back to run
    _fElapS := 0.0; // 作用域三：清衰减历时 / scope three, clear the decay duration
END_IF

// 段 3｜组态与输入域闸（R151 全覆盖）/ segment 3, the configuration and input domain gates
_bInOk := (iP = iP) AND ((iP - iP) = (iP - iP)) AND (iN = iN) AND ((iN - iN) = (iN - iN)); // 两电流有限性 / finiteness of both currents
_bCfgOk := (fBalLim > 0.0) AND (fBalLim = fBalLim) AND (fHystPct >= 0.0) AND (fHystPct <= fBalLim) AND (fStepThresh > 0.0) AND (fStepThresh = fStepThresh) AND (tDecayMax > T#0S) AND (fDtS > 0.0) AND (fDtS = fDtS); // 组态参数域判定 / the configuration domain verdict
IF (NOT _bInOk) OR (NOT _bCfgOk) OR ((ABS(iP) < 1.0E-6) AND (ABS(iN) < 1.0E-6)) THEN // 非有限、组态非法或双低电流（未出风）/ non finite, illegal config or both currents void
    IF NOT _bBad THEN // 未锁存才置 / set only while unlatched
        _bBad := TRUE; // 置传感器无效锁存 / raise the sensor bad latch
    END_IF
END_IF

// 段 4｜本拍平衡偏差计算（组合量）/ segment 4, the per scan balance deviation
_fDen := ABS(iP) + ABS(iN); // 电流幅值和 / the sum of magnitudes
IF _fDen > 1.0E-6 THEN // 幅值和可用 / the sum is usable
    _fDev := (iP - iN) / _fDen * 100.0; // 平衡偏差百分比，除子已证超阈 / the balance deviation with a proven divisor
ELSE // 幅值和不可用 / the sum is not usable
    _fDev := 0.0; // 偏差记零 / the deviation is zeroed
END_IF
fBalDevPct := _fDev; // 偏差出口 / the deviation outlet

// 段 5｜相位机：ENUM + CASE，含 ELSE 非法相位兜底（R128）/ segment 5, the phase machine with an ELSE fallback
CASE _ePhase OF
E_DL_VibPhase.eIdle: // 未使能相 / the disabled phase
    IF bEnable AND (NOT _bFault) THEN // 使能且无故障 / enabled and unfaulted
        _ePhase := E_DL_VibPhase.eRun; // 迁运行相 / migrate to run
    END_IF

E_DL_VibPhase.eRun: // 运行相：逐拍判级 + 步进突变检测 / the run phase, grading and the step detection
    IF NOT bEnable THEN // 失能 / disabled
        _ePhase := E_DL_VibPhase.eIdle; // 迁未使能相 / migrate to idle
    ELSIF _bBad THEN // 传感器无效锁存优先 / the sensor bad latch takes priority
        _bFault := TRUE; // 置故障锁存 / raise the fault latch
        _eFaulC := E_DL_VibFault.eSensorBad; // 故障级成因（R45 配对 bError）/ the fault cause paired with bError
        _ePhase := E_DL_VibPhase.eFault; // 迁故障相 / migrate to the fault phase
    ELSE // 正常判级 / the normal grading
        IF ABS(iP - _fIPrev) > fStepThresh THEN // 步进突变，起衰减测试 / a step change starts the decay test
            _fElapS := 0.0; // 历时清零 / clear the duration
            _ePhase := E_DL_VibPhase.eDecay; // 迁衰减相 / migrate to the decay phase
        END_IF
        IF _fDev > fBalLim THEN // 正偏进入判据 / the positive skew entry criterion
            _bPosL := TRUE; // 置正偏迟滞 / raise the positive latch
        ELSIF _fDev < fBalLim - fHystPct THEN // 正偏退出判据（迟滞收窄）/ the positive exit criterion
            _bPosL := FALSE; // 清正偏迟滞 / clear the positive latch
        END_IF
        IF _fDev < -fBalLim THEN // 负偏进入判据 / the negative skew entry criterion
            _bNegL := TRUE; // 置负偏迟滞 / raise the negative latch
        ELSIF _fDev > -fBalLim + fHystPct THEN // 负偏退出判据（迟滞收窄）/ the negative exit criterion
            _bNegL := FALSE; // 清负偏迟滞 / clear the negative latch
        END_IF
        bBalanced := (NOT _bPosL) AND (NOT _bNegL); // 平衡输出（迟滞派生）/ the balance outlet derived from the latches
        IF _bPosL THEN // 正偏故障（R190 独立成因）/ the positive skew fault, an independent cause
            _bFault := TRUE; // 置故障锁存 / raise the fault latch
            _eFaulC := E_DL_VibFault.ePosSkew; // 故障级成因（R45 配对 bError）/ the fault cause paired with bError
            _ePhase := E_DL_VibPhase.eFault; // 迁故障相 / migrate to the fault phase
        ELSIF _bNegL THEN // 负偏故障（R190 独立成因）/ the negative skew fault, an independent cause
            _bFault := TRUE; // 置故障锁存 / raise the fault latch
            _eFaulC := E_DL_VibFault.eNegSkew; // 故障级成因（R45 配对 bError）/ the fault cause paired with bError
            _ePhase := E_DL_VibPhase.eFault; // 迁故障相 / migrate to the fault phase
        END_IF
        _fIPrev := iP; // 快照推进 / advance the snapshot
    END_IF

E_DL_VibPhase.eDecay: // 衰减测试相：计时等待回带（退出条件 ≥2：回带 / 超时 / 失能，R98）/ the decay phase with at least two exit conditions
    IF NOT bEnable THEN // 失能 / disabled
        _ePhase := E_DL_VibPhase.eIdle; // 迁未使能相 / migrate to idle
    ELSIF _bBad THEN // 传感器无效 / the sensor went bad
        _bFault := TRUE; // 置故障锁存 / raise the fault latch
        _eFaulC := E_DL_VibFault.eSensorBad; // 故障级成因（R45 配对 bError）/ the fault cause paired with bError
        _ePhase := E_DL_VibPhase.eFault; // 迁故障相 / migrate to the fault phase
    ELSE // 计时中 / timing
        _fElapS := _fElapS + fDtS; // 历时累加 / accumulate the duration
        IF ABS(_fDev) <= fBalLim - fHystPct THEN // 偏差回带内（收窄带口径）/ the deviation is back inside the narrowed band
            fDecayS := _fElapS; // 衰减历时锁存 / latch the decay duration
            _ePhase := E_DL_VibPhase.eRun; // 迁回运行相 / migrate back to run
        ELSIF tonDecay.Q THEN // 衰减超时 / the decay timed out
            _bFault := TRUE; // 置故障锁存 / raise the fault latch
            _eFaulC := E_DL_VibFault.eDecaySlow; // 故障级成因（R45 配对 bError）/ the fault cause paired with bError
            _ePhase := E_DL_VibPhase.eFault; // 迁故障相 / migrate to the fault phase
        END_IF
        _fIPrev := iP; // 快照推进 / advance the snapshot
    END_IF

E_DL_VibPhase.eFault: // 故障相：成因锁存，等待复位沿 / the fault phase, the cause is latched until the reset edge
    IF NOT bEnable THEN // 失能 / disabled
        _ePhase := E_DL_VibPhase.eIdle; // 迁未使能相 / migrate to idle
    END_IF

ELSE // 非法相位兜底（R128）/ the illegal phase fallback
    _bFault := TRUE; // 置故障锁存 / raise the fault latch
    _eFaulC := E_DL_VibFault.ePhaseBad; // 故障级成因（R45 配对 bError）/ the fault cause paired with bError
    _ePhase := E_DL_VibPhase.eFault; // 迁故障相 / migrate to the fault phase
END_CASE

// 段 6｜统一出口 / segment 6, the unified outlet
IF _bFault THEN // 故障锁存优先 / the fault latch takes priority
    eFault := _eFaulC; // 故障级成因锁存回放（R152）/ the fault cause replayed from the latch
ELSE
    eFault := E_DL_VibFault.eNone; // 无锁存即无成因 / no latch, no cause
END_IF
ePhase := _ePhase; // 相位出口单点映射 / single point phase outlet mapping
bError := _bFault; // 故障标志与锁存位同源 / the fault flag shares the latch source
END_FUNCTION_BLOCK
